(* IEC 61131-3 sources: daoli-st-library/DL_Device (part 4) *)

(* ---- FB_DL_PortDiagAggregator.st ---- *)
(*==============================================================================
 * 组件名称 (Component)  : FB_DL_PortDiagAggregator
 * 所属子库 (Sublibrary) : DL_Device
 * 当前版本 (Version)    : 1.0.0
 * 组件分类 (Category)   : 功能块（FUNCTION_BLOCK）· 设备诊断 · 端口级聚合仲裁
 * 兼容性   (Platform)   : CODESYS 3.5 / TwinCAT 3 / 汇川 InoProShop / Schneider
 *                         Machine Expert；仅位与运算、TON、R_TRIG 与标准类型
 * 功能描述 (Function)   : 把最多 8 个现场总线通讯端口的链路状态、诊断码、
 *                         CRC 错误累计计数聚合成单一故障掩码、首出端口号、
 *                         首出诊断码与错误风暴标志，解决「多端口同时报警时
 *                         HMI 只看到最后一条」的现场痛点。本块只做端口级
 *                         （通讯物理端口）聚合与首出仲裁，不做模块级位域解析。
 * 边界声明 (Boundary)   : FB_DL_AxiolineDiagLatch 负责本地总线模块级（槽号加
 *                         位域）诊断锁存；FB_DL_PdiReadScheduler 负责参数对象
 *                         读取调度；本块数据源是「端口计数与端口诊断码」，
 *                         三者数据源不同、码段不共享、互不可替。
 * 首出语义 (First-out)  : 仅在无锁存时仲裁，同拍多端口故障取端口号最小者
 *                         （低号端口更靠近主站，是现场排故的默认因果顺序）；
 *                         锁存后不再更新，只有复位上升沿可清。复位处理放在
 *                         仲裁之后，保证复位当拍首出即为空，下一拍重新仲裁。
 * 拍序纪律 (Cycle order) : 本块属监视型，但「窗口差分」有硬拍序：增量必须在
 *                         装载前算出并转出，否则窗口结束拍装载当拍增量恒为 0。
 *                         故输出数组先转出（上一段快照）后装载（下一段基准）。
 * 风暴语义 (Burst)      : 风暴是趋势事件，不锁存；eBurst 只停留一拍，该拍
 *                         置 bBurstDetected 单拍标志，供上层做趋势记录或
 *                         降低总线负载，不参与 bError 判定。
 * 开源溯源 (Origin)     : plcnext-community / profibus-diag / namur-ne107。参考
 *                         PLCnext 官方帮助与 PROFIBUS 诊断公开手册的端口诊断
 *                         功能分类与参数域（端口号、链路状态、诊断码、错误
 *                         计数器、错误风暴阈值），只借分类与参数域，端口数
 *                         上限、掩码位序、枚举、状态机、码位与全部算法 100%
 *                         自有，输入一律经引脚注入，不绑定任何厂商系统变量，
 *                         clean-room 实现，不构成衍生作品。
 * 依赖     (Depends)    : 无 DL_ 内部依赖；仅 Standard.library 的 TON / R_TRIG
 * 故障码表 (Error codes):
 *   16#0003_0140【信息级】端口数超上限已钳位（只进码与趋势，不置故障位）
 *   16#0003_0141【信息级】统计窗口参数越界已钳位（只进码，不置故障位）
 *   16#0003_0300【故障级】端口故障锁存（伴随故障掩码非零，置 bError）
 *   16#0003_0301【故障级】诊断源未注入（端口数小于 1，置 bError）
 *   16#0003_0307【故障级】非法状态兜底（置 bError）
 * 码位占用 (Slot)       : 信息级 0140 / 0141；故障级 0300 / 0301 / 0307。
 *                         全部落在 R11 本件分配块内，无跨块借用。
 * 写入点次序 (Write order) :
 *   ① ePhase   ：段 8 状态机（唯一位移点），段 10 复位分支可回 eIdle
 *   ② uErrorId ：段 11 单一优先级链（0307 优于 0301 优于 0300 优于 0141
 *                 优于 0140），全拍只写一次，杜绝多分支互相覆盖
 *   ③ 首出锁存 ：段 9 仲裁（仅未锁存时）→ 段 10 复位（唯一清除点）
 *   ④ 基准计数 ：段 8 窗口结束拍装载，段 5 只读，永不与增量同拍混用
 * 验收向量 (Acceptance) :
 *   V1 端口 2 与端口 5 故障，其余正常 → 故障掩码 16#0012、存在端口故障为真
 *   V2 端口 5 先故障、端口 2 后故障 → 首出端口 5；复位后才可更新为 2
 *   V3 窗口 1 秒、阈值 10、端口 3 计数 100 增至 115 → 窗口结束拍增量为 15、
 *      风暴标志单拍为真
 *   V4 端口 4 计数 16#FFFF_FFFF 回绕到 3 → 增量为 3，不出现巨大正数
 *   V5 端口数 12 → 钳位 8、码 16#0003_0140、bError 为假
 * 红线自检 (Redline)    : R1 零全局变量表与外部变量引用 ｜ R2 零物理地址直写
 *                         R3 纯 IEC 61131-3 ｜ R4 防除零、防越界、无浮点判等
 *                         R5 全变量中英双语同行注释 ｜ R6 ENUM 加 CASE 加 ELSE
 *                         R7 TON 与 R_TRIG 全部在 CASE 之外无条件刷新
 *                         R8 信息级码不置 bError，故障级码才置
 * 修订历史 (Revision)   :
 *   2026-11-15  v1.0.0  首版落盘（Round 11 · 泳道 B · T1-7 端口诊断族）
 *============================================================================*)

(*------------------------------------------------------------------------------
 * 枚举: E_DL_PortDiagPhase（本块相位，归属本功能块并同文件发布）
 *       Phase enumeration owned by this block and published in the same file
 *-----------------------------------------------------------------------------*)
TYPE E_DL_PortDiagPhase :
(
    eIdle    := 0,   // 待机：未使能或端口数非法，掩码清零、首出保持 / Idle, mask cleared, first-out kept
    eMonitor := 10,  // 监视：逐拍算增量、逐端口去抖、窗口边界拍评估 / Monitoring, deltas and debounce running
    eBurst   := 20,  // 风暴：仅停留一拍，置单拍风暴标志后回监视 / Burst, one cycle only then back to monitor
    eFault   := 99   // 故障：诊断源缺失或非法状态，需复位退出 / Fault, needs a reset to leave
);
END_TYPE

(*------------------------------------------------------------------------------
 * 结构体: ST_DL_PortDiagState（跨周期状态，由调用方持有）
 *         Persistent state structure, owned by the caller
 *         注意：本结构体是跨周期数据，E_DL_PortDiagPhase 是相位枚举，
 *         二者刻意同名不同前缀，禁止相互替换使用
 *-----------------------------------------------------------------------------*)
TYPE ST_DL_PortDiagState :
STRUCT
    auPrevCnt   : ARRAY[1..8] OF UDINT;  // 上窗口各端口 CRC 计数基准 [次] / Previous window CRC counter per port
    nLatchPort  : INT;                   // 首出故障端口号 [1..8]，0 表示无 / First-out port number, zero means none
    uLatchCode  : UDINT;                 // 首出端口诊断码 [代码]，0 表示无 / First-out diagnostic code, zero means none
    bLatchValid : BOOL;                  // 首出锁存有效，仅复位可清 [-] / First-out latch valid, reset clears it
END_STRUCT
END_TYPE

(*==============================================================================
 * 逐拍推演 (Cycle-by-cycle trace)：
 *   场景 A 双端口故障（端口 2 与端口 5）
 *     拍 k 段 6 逐端口判定为真并启动各自去抖；段 9 见无锁存，取最小号端口 2
 *          锁存端口 2 与端口 2 的诊断码；段 11 掩码为 16#0012、置 0300
 *   场景 B 首出不覆盖（端口 5 先、端口 2 后）
 *     拍 k 端口 5 故障，锁存 5；拍 k+n 端口 2 也故障，但 bLatchValid 已真，
 *          段 9 只观测不覆盖，首出维持 5；复位后下一拍重新仲裁得 2
 *   场景 C 错误风暴（窗口 1 秒、阈值 10、端口 3 计数 100 增到 115）
 *     窗口内段 5 每拍算 115 减 100 得增量 15；窗口结束拍段 8 评估 15 大于 10，
 *          转 eBurst；下一拍 eBurst 置风暴单拍标志，回 eMonitor，同时已装载
 *          新基准 115，故下一窗口增量从 0 起算
 *   场景 D 计数回绕（端口 4 由 16#FFFF_FFFF 变为 3）
 *     段 5 判出当前值小于基准，按归零处理取 3，绝不出现巨大正数假风暴
 *   场景 E 端口数超上限（端口数 12）
 *     段 3 钳位为 8 并标记；段 11 单独置 0140，bError 保持假
 *============================================================================*)

FUNCTION_BLOCK FB_DL_PortDiagAggregator
VAR_INPUT
    bEnable          : BOOL;                              // 使能，FALSE 时掩码清零、首出保持 [-] / Enable, clears mask, holds first-out
    bReset           : BOOL;                              // 复位首出锁存，上升沿有效 [-] / Reset the first-out latch on a rising edge
    nPortCount       : INT;                               // 实际端口数 [个]，有效域 1 到 8 / Port count, valid range one to eight
    abPortLinkOk     : ARRAY[1..8] OF BOOL;               // 各端口链路正常标志 [TRUE=正常] / Per-port link up flags
    auPortErrCode    : ARRAY[1..8] OF UDINT;              // 各端口诊断码 [代码]，0 表示正常 / Per-port diagnostic code, zero means OK
    auPortCrcErrCnt  : ARRAY[1..8] OF UDINT;              // 各端口 CRC 错误累计计数 [次] / Per-port CRC error counter
    nBurstThreshold  : UDINT := 10;                       // 窗口内错误增量阈值 [次]，0 表示不判风暴 / Burst threshold per window, zero disables
    tBurstWindow     : TIME := T#1S;                      // 错误风暴统计窗口长度 [毫秒] / Burst evaluation window
    tDebounce        : TIME := T#200MS;                   // 端口故障确认去抖时间 [毫秒]，0 表示不去抖 / Port fault debounce, zero disables
END_VAR
VAR_OUTPUT
    bAnyPortFault    : BOOL;                              // 任一端口故障，等价掩码非零 [-] / Any port faulted, mask is non-zero
    bBurstDetected   : BOOL;                              // 错误风暴单拍标志，仅 eBurst 拍为真 [-] / Burst single-scan flag, true only in the burst cycle
    uPortFaultMask   : WORD;                              // 端口故障掩码，位 n 对应端口 n 加一 [位串] / Port fault mask, bit n is port n plus one
    nFirstFaultPort  : INT;                               // 首出故障端口号 [1..8]，0 表示无 / First-fault port number, zero means none
    uFirstFaultCode  : UDINT;                             // 首出端口诊断码 [代码]，与端口号同拍锁存 / First-fault diagnostic code latched with the port
    auPortDelta      : ARRAY[1..8] OF UDINT;              // 本窗口各端口错误增量 [次] / Per-port error increment of this window
    eState           : E_DL_PortDiagPhase;                // 主状态机当前相位 [-] / Current phase of the main state machine
    bError           : BOOL;                              // 故障级锁存，仅 0300 0301 0307 置位 [-] / Latched fault, only fault level codes set it
    uErrorId         : UDINT;                             // 事件码，0 表示无事件 [代码] / Event code, zero means none
END_VAR
VAR_IN_OUT
    stState          : ST_DL_PortDiagState;               // 跨周期状态：基准计数与首出锁存 [-] / Persistent state, baseline counters and first-out latch
END_VAR
VAR
    fbTrigReset      : R_TRIG;                            // 复位沿检测，CASE 之外无条件刷新 [-] / Reset edge detector, refreshed outside the CASE
    fbTonWindow      : TON;                               // 风暴统计窗口计时，CASE 之外无条件刷新 / Burst window timer, refreshed outside the CASE
    afbDebounce      : ARRAY[1..8] OF TON;                // 逐端口故障去抖定时器组，循环内无条件全刷新 / Per-port debounce timers, all refreshed every cycle
    bInit            : BOOL := FALSE;                     // 首扫标志，初值 FALSE，判据 NOT bInit [-] / First-scan flag initialised FALSE
    ePhase           : E_DL_PortDiagPhase := E_DL_PortDiagPhase.eIdle;  // 内部相位，对外经 eState 输出 / Internal phase, exported as eState
    nPortClamped     : INT;                               // 钳位后的端口数 [个]，0 到 8 / Clamped port count, zero to eight
    tWinUse          : TIME;                              // 实际生效的窗口长度 [毫秒] / Effective window length
    tDebUse          : TIME;                              // 实际生效的去抖时间 [毫秒] / Effective debounce time
    bWinRun          : BOOL;                              // 窗口计时器输入，边界拍拉低以重启窗口 / Window timer input, dropped on the boundary cycle
    bWinElapsed      : BOOL;                              // 窗口结束拍标志 [-] / Window boundary flag
    abRawFault       : ARRAY[1..8] OF BOOL;               // 端口原始故障（未去抖）[-] / Raw per-port fault before debouncing
    uMaskBuild       : WORD;                              // 去抖后故障掩码装配中间量 [位串] / Fault mask under assembly after debounce
    auRawDelta       : ARRAY[1..8] OF UDINT;              // 本拍增量装配中间量 [次] / Increment under assembly of this cycle
    auOutDelta       : ARRAY[1..8] OF UDINT;              // 增量输出快照，先转出后装载 [-] / Increment snapshot exported before reloading the baseline
    uMaxDelta        : UDINT;                             // 窗口内最大增量 [次] / Maximum increment inside the window
    nFirstScanPort   : INT;                               // 仲裁临时：最小号故障端口 [1..8] / Arbitration temporary, lowest faulted port
    uFirstScanCode   : UDINT;                             // 仲裁临时：该端口诊断码 [代码] / Arbitration temporary, that port diagnostic code
    bPortCntClamped  : BOOL;                              // 端口数超上限被钳位的标记 [-] / Flag, port count was clamped
    bParamClamped    : BOOL;                              // 时间参数越界被钳位的标记 [-] / Flag, a time parameter was clamped
    bStateIllegal    : BOOL;                              // 非法状态被兜底捕获的标记 [-] / Flag, an illegal state was captured
    i                : INT;                               // 端口遍历索引 [1..8] / Port loop index
END_VAR
VAR CONSTANT
    DL_PORT_MAX      : INT := 8;                          // 端口上限 [个] / Maximum port count
    DL_PORT_MASK_ALL : WORD := 16#00FF;                   // 八端口全掩码 [位串] / All eight port mask
    DL_MASK_ONE      : WORD := 16#0001;                   // 单端口基准位 [位串] / Single port base bit
    DL_WIN_MIN       : TIME := T#1MS;                     // 窗口长度下限 [毫秒]，防 0 窗口 / Minimum window length, guards a zero window
    DL_DEB_MIN       : TIME := T#1MS;                     // 去抖时间下限 [毫秒]，非零时套用 / Minimum debounce when not disabled
    DL_TIME_ZERO     : TIME := T#0MS;                     // 时间零值基准 [毫秒] / Time zero reference
    DL_BURST_MARGIN  : UDINT := 0;                        // 增量比较余量 [次]，保留语义位 / Increment comparison margin, reserved semantic slot
END_VAR

(*------------------------------------------------------------------------------
 * 段 1｜沿检测无条件刷新（R7 红线：CASE 之外每拍必刷）
 *      Edge detection refreshed unconditionally outside the CASE
 *-----------------------------------------------------------------------------*)
fbTrigReset(CLK := bReset);

(*------------------------------------------------------------------------------
 * 段 2｜首扫初始化（R19 唯一合法范式：初值 FALSE，判据 NOT bInit）
 *      First-scan initialisation, the canonical R19 pattern
 *-----------------------------------------------------------------------------*)
IF NOT bInit THEN
    FOR i := 1 TO DL_PORT_MAX DO
        stState.auPrevCnt[i] := 0;               // 基准计数清零，避免首窗口假风暴
        auOutDelta[i]        := 0;               // 增量输出清零，HMI 初值确定
    END_FOR
    stState.nLatchPort     := 0;                 // 首出端口号：0 表示无
    stState.uLatchCode     := 0;                 // 首出诊断码：0 表示无
    stState.bLatchValid    := FALSE;             // 首出锁存无效
    ePhase                 := E_DL_PortDiagPhase.eIdle;
    nPortClamped           := 0;
    uMaskBuild             := 16#0000;
    bWinRun                := FALSE;
    bBurstDetected         := FALSE;
    bPortCntClamped        := FALSE;
    bParamClamped          := FALSE;
    bStateIllegal          := FALSE;
    eState                 := E_DL_PortDiagPhase.eIdle;
    uErrorId               := 16#0000_0000;
    bError                 := FALSE;
    bInit                  := TRUE;              // 首扫只做一次
END_IF

(*------------------------------------------------------------------------------
 * 段 3｜端口数钳位（越界只钳位，不越界访问数组）
 *      Port count clamping, never index outside the array
 *-----------------------------------------------------------------------------*)
bPortCntClamped := FALSE;                        // 本拍标记预清零，避免历史残留
IF nPortCount < 1 THEN
    nPortClamped := 0;                           // 无诊断源：交由状态机转故障
ELSIF nPortCount > DL_PORT_MAX THEN
    nPortClamped    := DL_PORT_MAX;              // 超上限钳位到 8
    bPortCntClamped := TRUE;                     // 标记待置信息级码 0140
ELSE
    nPortClamped := nPortCount;
END_IF

(*------------------------------------------------------------------------------
 * 段 4｜时间参数钳位（0 有明确语义，不得与越界混为一谈）
 *      Time parameter clamping, zero keeps its documented meaning
 *-----------------------------------------------------------------------------*)
bParamClamped := FALSE;                          // 本拍标记预清零，避免历史残留
IF tBurstWindow <= DL_TIME_ZERO THEN
    tWinUse      := DL_WIN_MIN;                  // 0 窗口会让计时器每拍立即到期
    bParamClamped := TRUE;
ELSIF tBurstWindow < DL_WIN_MIN THEN
    tWinUse      := DL_WIN_MIN;
    bParamClamped := TRUE;
ELSE
    tWinUse := tBurstWindow;
END_IF

IF tDebounce < DL_TIME_ZERO THEN
    tDebUse      := DL_DEB_MIN;                  // 负时间不可能，按最小值兜底
    bParamClamped := TRUE;
ELSE
    tDebUse := tDebounce;                        // 0 表示不去抖，原样透传
END_IF

(*------------------------------------------------------------------------------
 * 段 5｜增量差分（回绕按归零处理，UDINT 语义不产生负数）
 *      Increment differencing, a wrapped counter is treated as a restart
 *      纪律：本段只读基准，装载基准只在段 8 窗口结束拍执行
 *-----------------------------------------------------------------------------*)
FOR i := 1 TO DL_PORT_MAX DO
    IF i > nPortClamped THEN
        auRawDelta[i] := 0;                      // 超出实际端口数一律记为 0
        auOutDelta[i] := 0;
    ELSIF auPortCrcErrCnt[i] < stState.auPrevCnt[i] THEN
        auRawDelta[i] := auPortCrcErrCnt[i];     // 计数器回绕或复位：按归零处理
        auOutDelta[i] := auRawDelta[i];
    ELSE
        auRawDelta[i] := auPortCrcErrCnt[i] - stState.auPrevCnt[i];
        auOutDelta[i] := auRawDelta[i];          // 先转出快照，供段 11 输出
    END_IF
END_FOR

(*------------------------------------------------------------------------------
 * 段 6｜端口故障判定与逐端口去抖（掩码装配）
 *      Per-port fault evaluation with per-port debounce and mask assembly
 *      定时器组在循环内对全部八端口无条件刷新，不因端口数少而漏刷
 *-----------------------------------------------------------------------------*)
uMaskBuild := 16#0000;
FOR i := 1 TO DL_PORT_MAX DO
    IF bEnable AND (i <= nPortClamped) AND ((NOT abPortLinkOk[i]) OR (auPortErrCode[i] <> UDINT#0)) THEN
        abRawFault[i] := TRUE;                   // 链路断或诊断码非零即原始故障
    ELSE
        abRawFault[i] := FALSE;
    END_IF
    afbDebounce[i](IN := abRawFault[i], PT := tDebUse);
    IF afbDebounce[i].Q THEN
        uMaskBuild := uMaskBuild OR SHL(DL_MASK_ONE, i - 1);  // 去抖成立才进位
    END_IF
END_FOR

(*------------------------------------------------------------------------------
 * 段 7｜窗口计时（无条件刷新，输入取自上一拍的运行允许位）
 *      Window timer refreshed unconditionally, input from the previous cycle
 *-----------------------------------------------------------------------------*)
fbTonWindow(IN := bWinRun, PT := tWinUse);
bWinElapsed := fbTonWindow.Q;

(*------------------------------------------------------------------------------
 * 段 8｜主状态机（ENUM 加 CASE，含 ELSE 兜底；每成员均有对应标签）
 *      Main state machine, one label per enumeration member plus a fallback
 *-----------------------------------------------------------------------------*)
bBurstDetected := FALSE;                         // 单拍标志预清零：只在 eBurst 拍置真
CASE ePhase OF
    E_DL_PortDiagPhase.eIdle:
        bWinRun := FALSE;                        // 待机不跑窗口，避免脏计时
        IF bEnable AND (nPortClamped >= 1) THEN
            ePhase  := E_DL_PortDiagPhase.eMonitor;
            bWinRun := TRUE;                     // 进入监视即启动首个窗口
        ELSIF bEnable AND (nPortClamped < 1) THEN
            ePhase := E_DL_PortDiagPhase.eFault; // 诊断源未注入：故障级 0301
        END_IF

    E_DL_PortDiagPhase.eMonitor:
        IF NOT bEnable THEN
            ePhase     := E_DL_PortDiagPhase.eIdle;
            bWinRun    := FALSE;
            uMaskBuild := 16#0000;               // 未使能掩码清零，首出保持
        ELSIF nPortClamped < 1 THEN
            ePhase  := E_DL_PortDiagPhase.eFault;
            bWinRun := FALSE;
        ELSIF bWinElapsed THEN
            uMaxDelta     := 0;                  // 窗口结束拍：求最大增量
            FOR i := 1 TO nPortClamped DO
                IF auRawDelta[i] > uMaxDelta THEN
                    uMaxDelta := auRawDelta[i];
                END_IF
            END_FOR
            IF (nBurstThreshold > UDINT#0) AND (uMaxDelta > (nBurstThreshold + DL_BURST_MARGIN)) THEN
                ePhase := E_DL_PortDiagPhase.eBurst;   // 超阈值：下一拍置单拍标志
            ELSE
                ePhase := E_DL_PortDiagPhase.eMonitor; // 未超阈值：原地自保持
            END_IF
            FOR i := 1 TO DL_PORT_MAX DO
                stState.auPrevCnt[i] := auPortCrcErrCnt[i];  // 装载新基准
            END_FOR
            bWinRun := FALSE;                    // 拉低一拍，强制窗口重新起算
        ELSE
            bWinRun := TRUE;                     // 窗口内持续计时
        END_IF

    E_DL_PortDiagPhase.eBurst:
        bBurstDetected := TRUE;                  // 仅此一拍为真，不锁存，不进故障
        bWinRun        := FALSE;                 // 风暴拍不重启窗口，下一拍再说
        ePhase         := E_DL_PortDiagPhase.eMonitor;

    E_DL_PortDiagPhase.eFault:
        uMaskBuild := 16#0000;                   // 故障态不外送掩码，防误联锁
        bWinRun    := FALSE;
        IF NOT bEnable THEN
            ePhase := E_DL_PortDiagPhase.eIdle;  // 停使能可直接退出故障态
        END_IF

    ELSE
        ePhase        := E_DL_PortDiagPhase.eFault;   // 非法值兜底
        uMaskBuild    := 16#0000;
        bWinRun       := FALSE;
        bStateIllegal := TRUE;                   // 由段 11 统一置 0307
END_CASE

(*------------------------------------------------------------------------------
 * 段 9｜首出仲裁（仅未锁存时执行；升序取最小号端口，先到先得）
 *      First-out arbitration, only when not yet latched, lowest port wins
 *-----------------------------------------------------------------------------*)
IF (NOT stState.bLatchValid) AND uMaskBuild <> 16#0000 THEN
    nFirstScanPort := 0;
    uFirstScanCode := 0;
    FOR i := 1 TO nPortClamped DO
        IF ((uMaskBuild AND SHL(DL_MASK_ONE, i - 1)) <> 16#0000) AND (nFirstScanPort = 0) THEN
            nFirstScanPort := i;                       // 升序首个命中即最小号端口
            uFirstScanCode := auPortErrCode[i];
        END_IF
    END_FOR
    IF nFirstScanPort > 0 THEN
        stState.nLatchPort  := nFirstScanPort;
        stState.uLatchCode  := uFirstScanCode;
        stState.bLatchValid := TRUE;                   // 锁存后本窗口不再改写
    END_IF
END_IF

(*------------------------------------------------------------------------------
 * 段 10｜复位（放在仲裁之后，保证复位当拍首出即为空）
 *      Reset placed after arbitration so the first-out is empty this cycle
 *-----------------------------------------------------------------------------*)
IF fbTrigReset.Q THEN
    stState.nLatchPort  := 0;
    stState.uLatchCode  := 0;
    stState.bLatchValid := FALSE;
    bError              := FALSE;
    bStateIllegal       := FALSE;
    ePhase              := E_DL_PortDiagPhase.eIdle;   // 复位后回待机，再按使能重入
    bWinRun             := FALSE;
END_IF

(*------------------------------------------------------------------------------
 * 段 11｜输出归并与码位定级（单一优先级链，全拍只写一次 uErrorId）
 *      Output merge and single-priority error code resolution
 *-----------------------------------------------------------------------------*)
uPortFaultMask  := uMaskBuild AND DL_PORT_MASK_ALL;    // 屏蔽高位脏数据
bAnyPortFault   := (uPortFaultMask <> 16#0000);
nFirstFaultPort := stState.nLatchPort;
uFirstFaultCode := stState.uLatchCode;

IF bStateIllegal THEN
    uErrorId := 16#0003_0307;                          // 优先级一：非法状态
ELSIF (nPortClamped < 1) AND bEnable THEN
    uErrorId := 16#0003_0301;                          // 优先级二：诊断源缺失
ELSIF uPortFaultMask <> 16#0000 THEN
    uErrorId := 16#0003_0300;                          // 优先级三：端口故障锁存
ELSIF bParamClamped THEN
    uErrorId := 16#0003_0141;                          // 信息级：参数越界已钳位
ELSIF bPortCntClamped THEN
    uErrorId := 16#0003_0140;                          // 信息级：端口数越界已钳位
ELSE
    uErrorId := 16#0000_0000;
END_IF

(* 故障位只反映故障级：信息级码 0140 与 0141 绝不置故障位（R21） *)
bError := bStateIllegal
          OR ((nPortClamped < 1) AND bEnable)
          OR (uPortFaultMask <> 16#0000);

eState          := ePhase;                             // 相位每拍重写，供 HMI 诊断
auPortDelta[1]  := auOutDelta[1];                      // 增量数组逐元素转出，避免整数组赋值
auPortDelta[2]  := auOutDelta[2];
auPortDelta[3]  := auOutDelta[3];
auPortDelta[4]  := auOutDelta[4];
auPortDelta[5]  := auOutDelta[5];
auPortDelta[6]  := auOutDelta[6];
auPortDelta[7]  := auOutDelta[7];
auPortDelta[8]  := auOutDelta[8];
END_FUNCTION_BLOCK

(* ---- FB_DL_PortDiagBoard.st ---- *)
(*==============================================================================
 * 组件名称 (Component)  : FB_DL_PortDiagBoard
 * 所属子库 (Sublibrary) : DL_Device
 * 当前版本 (Version)    : 1.0.0
 * 组件分类 (Category)   : 功能块（FUNCTION_BLOCK）· 设备诊断 · 多组端口看板与首出仲裁
 * 兼容性   (Platform)   : CODESYS 3.5 / TwinCAT 3 / 汇川 InoProShop / Schneider
 *                         Machine Expert；纯 IEC 61131-3（第 3 版）语法，
 *                         仅依赖 Standard.library（R_TRIG），零厂商方言
 * 功能描述 (Function)   : 把最多 4 个端口诊断聚合组（每组最多 8 端口）汇总为一张看板：
 *                         屏蔽超界位后的各组掩码、全局故障端口总数、全局首出端口
 *                         （组号加端口号加诊断码），以及按「组号优先、端口号次之」稳定
 *                         排序的前 3 个待修端口。回答现场两个问题：现在还剩几个端口坏、
 *                         先修哪一个。
 * 分层声明 (Layering)   : ① 本件是「汇总层」，只消费端口级聚合结果（掩码加组内首出
 *                         码），不实例化上游聚合块、不重算端口明细——聚合器实例由调用方
 *                         按组各自持有，重复实例化会造成同一批端口被算两遍；
 *                         ② 不读模块级状态字（模块级归本地总线诊断锁存件，端口级归聚合
 *                         器，参数对象级归参数回读调度件，三层数据源分账已在 R11 收口）；
 *                         ③ 不绑定任何总线驱动，全部数据经引脚注入。
 * 职责边界 (Scope)      : 不做端口去抖（聚合器职责）、不做报警确认与搁置、不做历史趋势
 *                         归档、不做跨机架分组切换（组数运行期变化按钳位处理）。
 * 组数语义 (Grouping)   : 组是「同一块远程 IO 卡或同一台交换机的 8 个端口」的物理分组，
 *                         组号小者更靠近主站，故首出仲裁取组号最小、再取端口号最小，
 *                         这与现场排故的因果顺序一致。
 * 开源溯源 (Origin)     : 来源标签 plcnext-diag 加 roadmap-p0。原创实现（参考 T1-7
 *                         PLCnext 端口诊断四元组的分类与参数域，以及 ROADMAP §15.3 P0
 *                         条目的「看板加首出」需求定义）。仅借分类层次、参数域与验收
 *                         口径，掩码位序、首出三律、Top 排序编码、枚举、状态机与全部
 *                         码位 100% 本库独立设计，clean-room 实现，零代码行复制。
 *                         PLCnext 帮助文档为厂商公开资料，此处按最严口径「只借结构与
 *                         参数域」处置，不构成衍生作品。
 * 依赖     (Depends)    : 无 DL_ 内部依赖；Standard.library: R_TRIG
 * 故障码表 (Error codes):
 *   16#0003_0149【信息级】组数超上限已钳位到 4（只影响显示范围，不置故障位）
 *   16#0003_014A【信息级】某组端口数超上限已钳位到 8（组态常见，非错误）
 *   16#0003_014B【信息级】掩码超界位已屏蔽（绝不把不存在的端口计入故障数）
 *   16#0003_014C【信息级】组内声明首出端口与掩码推导值不一致（数据源未同步）
 *   16#0003_030B【故障段趋势码】单拍掩码变化位数超阈值，判为组态刷新；按规格
 *                         第 3.13 节「仅提示不锁存」处置：只透出一拍，不置故障位
 *   16#0003_0309【故障级】组数小于 1，无诊断源（锁存，置故障位）
 *   16#0003_030A【故障级】某组端口数小于 1，该组掩码含义不可信（锁存，置故障位）
 *   16#0003_030C【故障级】非法状态兜底（锁存，置故障位，终端安全态）
 * 码位占用 (Slot)       : 信息级 0149 / 014A / 014B / 014C；故障级 0309 / 030A / 030B / 030C。
 *                         全部落在 R12 本件分配块内，无跨块借用、无段外哨兵值。
 * 拍序纪律 (Cycle order) :
 *   ① ePhase      ：段 4 状态机（唯一位移点），段 6 复位分支是唯一回退点
 *   ② 首出锁存    ：段 4 的 eScanning 分支（仅未锁存时仲裁）→ 段 5 换出 → 段 6 复位清除
 *   ③ 输出码      ：段 7 单一优先级链，全拍只写一次 uErrorId，杜绝多分支互相覆盖
 *   ④ 掩码基准    ：段 4 的 eScanning 分支末尾装载，与风暴判定同段且判在读后写前
 * 首出三律 (First-out)  : ① 仅在无锁存时仲裁；② 同拍多端口故障取组号最小、再取端口号
 *                         最小；③ 复位在仲裁之后执行，故复位当拍首出为空、下一拍重新
 *                         仲裁（与 R11 端口聚合器同口径）。
 * 验收向量 (Acceptance) :
 *   V1 单组超界位：组数 1、端口数 8、掩码 16#0101 → 位 8 对应端口 9 超界被屏蔽，
 *      掩码出 16#0001、总故障 1、首出 1 组 1 号、码 014B
 *   V2 双组排序：两组端口数 8，掩码 16#0004 与 16#0003 → 总数 3、首出 1 组 3 号、
 *      待修序 13、21、22（编码为组号乘 10 加端口号）
 *   V3 复位时序：与 V2 同参，复位上升沿当拍首出为空，下一拍重新仲裁回 1 组 3 号
 *   V4 无诊断源：组数 0 → 钳为 1、故障位置位、码 0309
 *   V5 空组：第 1 组端口数 0 → 钳为 1、故障位置位、码 030A
 * 偏离留档 (Deviation)  :
 *   ① 规格第 3.13 节算法要点对「端口数超上限」写 014A、对「端口数越界」的边界说明
 *      又写 030A。本件按语义拆分：大于 8 属组态多填，按信息级 014A 只钳位；小于 1
 *      属无有效端口（掩码含义不可信），按故障级 030A 锁存——与验收向量 V5 完全一致。
 *   ② 规格未给 anGroupFirstPort 的用途。本件把它用作「声明值与掩码推导值」的一致性
 *      校验（为 0 视为未填、不校验），不一致只置信息级 014C，避免该引脚悬空无意义。
 *   ③ 030B 落在故障段但不置故障位，理由见上方故障码表，属规格原文要求的「仅提示不
 *      锁存」，不是定级笔误。
 * 修订历史 (Revision)   :
 *   2026-11-15  v1.0.0  首版落盘（R12 · 泳道 C · 端口诊断看板 P0 件）
 *============================================================================*)

(*------------------------------------------------------------------------------
 * 枚举: E_DL_BoardPhase（本块相位，归属本功能块并同文件发布）
 *       Phase enumeration owned by this block and published in the same file
 *-----------------------------------------------------------------------------*)
TYPE E_DL_BoardPhase :
(
    eIdle     := 0,   // 待机：钳位参数后即转扫描，或未使能时清掩码保首出 / Idle, clamps parameters then moves on to scanning
    eScanning := 10,  // 扫描：一趟完成屏蔽、计数、首出仲裁与待修排序，本拍结束回待机 / Scanning, the whole sweep completes in one pass
    eFault    := 99   // 故障：无诊断源、空组或非法状态，需复位退出 / Fault, needs a reset to leave
);
END_TYPE

(*------------------------------------------------------------------------------
 * 结构体: ST_DL_BoardState（跨周期状态，由调用方持有）
 *         Persistent state structure, owned by the caller
 *         说明：首出锁存是「诊断证据」，掉使能不清、只有复位沿才清；
 *               anLastMask 用于掩码跳变风暴的差分基准
 *-----------------------------------------------------------------------------*)
TYPE ST_DL_BoardState :
STRUCT
    nLatchedGroup : INT;                     // 首出锁存组号 [1..4]，0 表示无 / Latched first-out group, zero means none
    nLatchedPort  : INT;                     // 首出锁存端口号 [1..8]，0 表示无 / Latched first-out port, zero means none
    uLatchedCode  : UDINT;                   // 首出锁存诊断码 [代码]，0 表示未填 / Latched first-out diagnostic code, zero means not filled
    bLatchValid   : BOOL;                    // 首出锁存有效，仅复位沿可清 / First-out latch valid, cleared by the reset edge only
    anLastMask    : ARRAY[1..4] OF WORD;     // 上次各组掩码快照，用于跳变风暴差分 [位串] / Previous per-group mask for burst differencing
END_STRUCT
END_TYPE

FUNCTION_BLOCK FB_DL_PortDiagBoard
VAR_INPUT
    bEnable          : BOOL;                              // 看板使能，FALSE 时掩码清零而首出保持 [-] / Enable, masks are cleared while the first-out latch is kept
    bReset           : BOOL;                              // 复位首出锁存，上升沿有效 [-] / Rising edge clears the first-out latch
    nGroupCount      : INT := 1;                          // 聚合组数 [组]，有效域 1 到 4 / Group count, valid range one to four
    anGroupFaultMask : ARRAY[1..4] OF WORD;               // 各组端口故障掩码，位 n 减一 对应端口 n [位串] / Per-group fault mask, bit n minus one is port n
    anGroupPortCount : ARRAY[1..4] OF INT;                // 各组实际端口数 [个]，有效域 1 到 8 / Ports per group, valid range one to eight
    anGroupFirstPort : ARRAY[1..4] OF INT;                // 各组声明首出端口号，0 表示未填不校验 [端口号] / Declared first-out port, zero skips the cross check
    auGroupFirstCode : ARRAY[1..4] OF UDINT;              // 各组组内首出诊断码 [代码]，0 表示未填 / Per-group first-out diagnostic code, zero means not filled
END_VAR
VAR_OUTPUT
    nTotalFaultPort  : INT;                               // 全局故障端口总数 [个] / Total faulted ports across the enabled groups
    nFirstGroup      : INT;                               // 全局首出组号 [1..4]，0 表示无 / Global first-out group, zero means none
    nFirstPort       : INT;                               // 全局首出端口号 [1..8]，0 表示无 / Global first-out port, zero means none
    uFirstCode       : UDINT;                             // 全局首出诊断码 [代码]，0 表示未填 / Global first-out diagnostic code
    anGroupMaskOut   : ARRAY[1..4] OF WORD;               // 屏蔽超界位后的各组掩码 [位串] / Sanitised per-group masks
    anTopPortNo      : ARRAY[1..3] OF INT;                // 待修端口编码，组号乘 10 加端口号，0 表示空位 [编码] / Top repair ports encoded as group times ten plus port
    auTopPortCode    : ARRAY[1..3] OF UDINT;              // 待修端口对应诊断码 [代码] / Diagnostic code of each top repair port
    bAnyFault        : BOOL;                              // 总故障数大于 0 [-] / Any faulted port present
    bError           : BOOL;                              // 故障级锁存，仅 0309 030A 030C 置位 [-] / Latched fault, only fault level codes set it
    uErrorId         : UDINT;                             // 事件码，0 表示无事件 [代码] / Event code, zero means none
    eState           : E_DL_BoardPhase;                   // 主状态机当前相位 [-] / Current phase of the main state machine
END_VAR
VAR_IN_OUT
    stBoard          : ST_DL_BoardState;                  // 跨周期：首出锁存与掩码差分基准 [-] / Persistent first-out latch and mask baseline
END_VAR
VAR
    fbTrigReset      : R_TRIG;                            // 复位沿检测，主周期无条件刷新 [-] / Reset edge detector, refreshed unconditionally
    ePhase           : E_DL_BoardPhase := E_DL_BoardPhase.eIdle; // 内部相位，对外经 eState 输出 [-] / Internal phase exported as eState
    bInit            : BOOL := FALSE;                     // 首扫标志，初值 FALSE，判据取非 [-] / First-scan flag initialised FALSE
    bMaskBase        : BOOL := FALSE;                     // 掩码差分基准已装载 [-] / Mask baseline loaded flag
    bFaultLatch      : BOOL;                              // 故障锁存，仅复位分支清除 [-] / Fault latch, cleared by the reset path only
    uErrInt          : UDINT;                             // 故障级码寄存，锁存型 [代码] / Latched fault level code register
    uInfoCode        : UDINT;                             // 本拍信息级码，每拍重算 [代码] / Info level code recomputed every scan
    nGroupUse        : INT;                               // 生效组数，钳位后 [组] / Effective group count after clamping
    auPortCntUse     : ARRAY[1..4] OF INT;                // 生效端口数，钳位后 [个] / Effective port count per group after clamping
    uBuildMask       : WORD;                              // 掩码装配中间量 [位串] / Mask under assembly
    uDiff            : WORD;                              // 掩码差分中间量 [位串] / Mask difference under evaluation
    nTotal           : INT;                               // 故障端口累加计数 [个] / Faulted port counter
    nMinPort         : INT;                               // 组内最小故障端口号 [1..8]，0 表示无 / Lowest faulted port inside a group
    nBitScan         : INT;                               // 掩码跳变位计数 [位] / Changed bit counter for the burst check
    nScanGroup       : INT;                               // 仲裁扫描组号 [1..4] / Arbitration group index
    nScanPort        : INT;                               // 仲裁扫描端口号 [1..8] / Arbitration port index
    bFound           : BOOL;                              // 仲裁命中标志 [-] / Arbitration hit flag
    nTopCount        : INT;                               // 已填待修位个数 [个] / Filled top repair slots
    nGuard           : DINT;                              // 循环守卫计数 [次]，上限常量化 / Loop guard counter with a constant bound
    bMaskClamped     : BOOL;                              // 本拍存在掩码超界位被屏蔽 [-] / Mask bits were suppressed this scan
    bPortClamped     : BOOL;                              // 本拍存在端口数超上限被钳位 [-] / A port count was clamped this scan
    bGroupClamped    : BOOL;                              // 本拍组数超上限被钳位 [-] / The group count was clamped this scan
    bPortShort       : BOOL;                              // 本拍存在某组端口数小于 1 [-] / A group has no usable port this scan
    bGroupShort      : BOOL;                              // 本拍组数小于 1 [-] / The group count is below one this scan
    bPortDeclMismatch: BOOL;                              // 声明首出端口与推导值不一致 [-] / Declared first-out port differs from the derived one
    bMaskJump        : BOOL;                              // 单拍掩码跳变位超阈值 [-] / Mask changed in more bits than the threshold
    g                : INT;                               // 组循环索引 [1..4] / Group loop index
    p                : INT;                               // 端口循环索引 [1..8] / Port loop index
END_VAR
VAR CONSTANT
    DL_GROUP_MAX     : INT := 4;                          // 聚合组数上限 [组] / Maximum group count
    DL_PORT_MAX      : INT := 8;                          // 组内端口数上限 [个] / Maximum ports per group
    DL_TOP_N         : INT := 3;                          // 待修输出位个数 [个] / Number of top repair slots
    DL_GROUP_STRIDE  : INT := 10;                         // 端口编码步长，组号乘该值加端口号 / Encoding stride of the top repair code
    DL_JUMP_MAX      : INT := 8;                          // 单拍掩码跳变位阈值 [位] / Changed bit threshold per scan
    DL_GUARD_MAX     : DINT := 96;                        // 循环守卫上限 [次] / Loop guard bound
    DL_WORD_BITS     : INT := 16;                         // 掩码字宽，超界位屏蔽的遍历上限 [位] / Mask word width
    DL_MASK_ONE      : WORD := 16#0001;                   // 单端口基准位 [位串] / Single port base bit
    DL_MASK_NONE     : WORD := 16#0000;                   // 全零掩码基准 [位串] / All zero mask reference
END_VAR

(*------------------------------------------------------------------------------
 * 段 1｜输出确定性默认值（公约：出口先赋；单拍标志每拍预清零，R25 第一律）
 *      Deterministic defaults first, one-scan flags pre-cleared every scan
 *-----------------------------------------------------------------------------*)
bAnyFault         := FALSE;                     // 看板派生量预清零（Dashboard flag pre-cleared）
uInfoCode         := 16#0000_0000;              // 信息级码每拍重算（Info code recomputed every scan）
bMaskClamped      := FALSE;                     // 掩码屏蔽标记预清零（Mask suppression flag pre-cleared）
bPortClamped      := FALSE;                     // 端口数钳位标记预清零（Port clamp flag pre-cleared）
bGroupClamped     := FALSE;                     // 组数钳位标记预清零（Group clamp flag pre-cleared）
bPortShort        := FALSE;                     // 空组标记预清零（Empty group flag pre-cleared）
bGroupShort       := FALSE;                     // 无组标记预清零（No group flag pre-cleared）
bPortDeclMismatch := FALSE;                     // 声明一致性标记预清零（Declared mismatch flag pre-cleared）
bMaskJump         := FALSE;                     // 掩码跳变标记预清零（Mask jump flag pre-cleared）
nGuard            := 0;                         // 循环守卫清零（Loop guard cleared）

(*------------------------------------------------------------------------------
 * 段 2｜沿检测无条件刷新（红线：实例在 CASE 之外每拍必刷）
 *      Edge detection refreshed unconditionally outside the CASE
 *-----------------------------------------------------------------------------*)
fbTrigReset(CLK := bReset);

(*------------------------------------------------------------------------------
 * 段 3｜首扫初始化（唯一合法范式：初值 FALSE，判据取非）
 *      First-scan initialisation following the single legal pattern
 *-----------------------------------------------------------------------------*)
IF NOT bInit THEN
    FOR g := 1 TO DL_GROUP_MAX DO
        stBoard.anLastMask[g] := DL_MASK_NONE;  // 掩码差分基准清零，避免首拍假风暴（Baseline cleared to suppress a false burst）
        anGroupMaskOut[g]     := DL_MASK_NONE;  // 掩码出口清零，HMI 初值确定（Mask outlet cleared for a deterministic HMI start value）
    END_FOR
    FOR p := 1 TO DL_TOP_N DO
        anTopPortNo[p]   := 0;                  // 待修端口空位（Top repair slot empty）
        auTopPortCode[p] := 0;                  // 待修诊断码清零（Top repair code cleared）
    END_FOR
    stBoard.nLatchedGroup := 0;                 // 首出组号：0 表示无（No first-out group）
    stBoard.nLatchedPort  := 0;                 // 首出端口号：0 表示无（No first-out port）
    stBoard.uLatchedCode  := 0;                 // 首出码：0 表示未填（No first-out code）
    stBoard.bLatchValid   := FALSE;             // 首出锁存无效（First-out latch invalid）
    nTotalFaultPort       := 0;                 // 故障总数清零（Fault total cleared）
    nFirstGroup           := 0;                 // 首出组号出口清零（First-out group outlet cleared）
    nFirstPort            := 0;                 // 首出端口出口清零（First-out port outlet cleared）
    uFirstCode            := 0;                 // 首出码出口清零（First-out code outlet cleared）
    bFaultLatch           := FALSE;             // 故障锁存清零（Fault latch cleared）
    uErrInt               := 16#0000_0000;      // 故障码清零（Fault code cleared）
    bMaskBase             := FALSE;             // 差分基准待本拍装载（Baseline to be loaded this scan）
    ePhase                := E_DL_BoardPhase.eIdle; // 相位复位为待机（Phase reset to idle）
    bInit                 := TRUE;              // 首扫只做一次（First scan runs once）
END_IF

(*------------------------------------------------------------------------------
 * 段 4｜主状态机（枚举每个成员均有标签，末尾 ELSE 兜底到终端安全态）
 *      Main state machine, one label per member plus a trailing ELSE fallback
 *-----------------------------------------------------------------------------*)
CASE ePhase OF

    E_DL_BoardPhase.eIdle: // 待机：未使能则清掩码保首出，使能则钳位参数后转扫描
        IF NOT bEnable THEN
            FOR g := 1 TO DL_GROUP_MAX DO
                anGroupMaskOut[g] := DL_MASK_NONE;  // 掉使能掩码清零，防止下游误联锁（Masks cleared while disabled）
            END_FOR
            nTotalFaultPort := 0;               // 故障总数清零（Fault total cleared）
            bAnyFault       := FALSE;           // 无故障派生量（No fault derived）
            ePhase          := E_DL_BoardPhase.eIdle; // 保持在待机（Stay idle）
        ELSE
            IF nGroupCount < 1 THEN
                nGroupUse    := 1;              // 无组：先给 1 供后续诊断（Fall back to one group）
                bGroupShort  := TRUE;           // 标记待置 0309（Flag for code 0309）
            ELSIF nGroupCount > DL_GROUP_MAX THEN
                nGroupUse    := DL_GROUP_MAX;   // 超上限钳位（Clamp to the upper bound）
                bGroupClamped := TRUE;          // 标记待置 0149（Flag for code 0149）
            ELSE
                nGroupUse := nGroupCount;       // 合法组数直通（Valid group count passed through）
            END_IF
            FOR g := 1 TO DL_GROUP_MAX DO
                nGuard := nGuard + 1;           // 守卫递增（Guard incremented）
                IF nGuard > DL_GUARD_MAX THEN
                    EXIT;                       // 守卫到顶即退出，防死循环（Bail out at the guard bound）
                END_IF
                IF g <= nGroupUse THEN
                    IF anGroupPortCount[g] < 1 THEN
                        auPortCntUse[g] := 1;   // 空组：先给 1 供后续诊断（Empty group falls back to one port）
                        bPortShort      := TRUE; // 标记待置 030A（Flag for code 030A）
                    ELSIF anGroupPortCount[g] > DL_PORT_MAX THEN
                        auPortCntUse[g] := DL_PORT_MAX; // 超上限钳位（Clamp to the upper bound）
                        bPortClamped    := TRUE;        // 标记待置 014A（Flag for code 014A）
                    ELSE
                        auPortCntUse[g] := anGroupPortCount[g]; // 合法端口数直通（Valid port count passed through）
                    END_IF
                ELSE
                    auPortCntUse[g] := 0;       // 未启用组记 0，不参与扫描（Unused group marked zero）
                END_IF
            END_FOR
            IF bGroupShort THEN
                bFaultLatch := TRUE;                        // 无诊断源：锁故障（No diagnostic source, latch a fault）
                uErrInt     := 16#0003_0309;                // 0309 组数小于 1（Group count below one）
                ePhase      := E_DL_BoardPhase.eFault;      // 进故障态（Enter the fault state）
            ELSIF bPortShort THEN
                bFaultLatch := TRUE;                        // 空组：锁故障（Empty group latches a fault）
                uErrInt     := 16#0003_030A;                // 030A 端口数小于 1（Port count below one）
                ePhase      := E_DL_BoardPhase.eFault;      // 进故障态（Enter the fault state）
            ELSE
                ePhase := E_DL_BoardPhase.eScanning;        // 参数可用，进入扫描（Parameters usable, start scanning）
            END_IF
        END_IF

    E_DL_BoardPhase.eScanning: // 扫描：屏蔽、计数、首出仲裁、待修排序、跳变差分，一趟完成
        nTotal    := 0;                         // 故障计数清零（Fault counter cleared）
        nBitScan  := 0;                         // 跳变位计数清零（Changed bit counter cleared）
        (* ① 屏蔽超界位并统计故障数，同时取组内最小故障端口号 *)
        nGuard := 0;                            // 子段守卫清零（Guard reset for this pass）
        FOR g := 1 TO DL_GROUP_MAX DO
            nGuard := nGuard + 1;               // 守卫递增（Guard incremented）
            IF nGuard > DL_GUARD_MAX THEN
                EXIT;                           // 守卫到顶即退出（Bail out at the guard bound）
            END_IF
            IF g <= nGroupUse THEN
                uBuildMask := anGroupFaultMask[g];      // 取原始掩码（Take the raw mask）
                nMinPort   := 0;                        // 组内最小端口号预清零（Lowest port pre-cleared）
                FOR p := 1 TO DL_WORD_BITS DO
                    nGuard := nGuard + 1;               // 守卫递增（Guard incremented）
                    IF nGuard > DL_GUARD_MAX THEN
                        EXIT;                           // 守卫到顶即退出（Bail out at the guard bound）
                    END_IF
                    IF p > auPortCntUse[g] THEN
                        IF (uBuildMask AND SHL(DL_MASK_ONE, p - 1)) <> DL_MASK_NONE THEN
                            bMaskClamped := TRUE;       // 超界位有值：标记待置 014B（Out-of-range bit held a value）
                        END_IF
                        uBuildMask := uBuildMask AND (NOT SHL(DL_MASK_ONE, p - 1)); // 超界位清零（Clear the out-of-range bit）
                    ELSE
                        IF (uBuildMask AND SHL(DL_MASK_ONE, p - 1)) <> DL_MASK_NONE THEN
                            nTotal := nTotal + 1;       // 在界内且为故障：计数（In range and faulted, count it）
                            IF nMinPort = 0 THEN
                                nMinPort := p;          // 首次命中即组内最小号（First hit is the lowest port）
                            END_IF
                        END_IF
                    END_IF
                END_FOR
                anGroupMaskOut[g] := uBuildMask;        // 屏蔽后掩码出口（Sanitised mask outlet）
                IF (anGroupFirstPort[g] > 0) AND (anGroupFirstPort[g] <> nMinPort) THEN
                    bPortDeclMismatch := TRUE;          // 声明值与推导值不一致：标记 014C（Declared value differs, flag 014C）
                END_IF
            ELSE
                anGroupMaskOut[g] := DL_MASK_NONE;      // 未启用组掩码清零（Unused group mask cleared）
            END_IF
        END_FOR
        nTotalFaultPort := nTotal;              // 故障总数出口（Fault total outlet）
        bAnyFault       := (nTotal > 0);        // 存在故障（Any fault present）
        (* ② 首出仲裁：仅未锁存时执行，组号优先、端口号次之，取字典序最小 *)
        nGuard := 0;                            // 子段守卫清零（Guard reset for this pass）
        IF (NOT stBoard.bLatchValid) AND (nTotal > 0) THEN
            bFound      := FALSE;               // 命中标志预清零（Hit flag pre-cleared）
            nScanGroup  := 0;                   // 仲裁组号预清零（Arbitration group pre-cleared）
            nScanPort   := 0;                   // 仲裁端口号预清零（Arbitration port pre-cleared）
            FOR g := 1 TO nGroupUse DO
                nGuard := nGuard + 1;           // 守卫递增（Guard incremented）
                IF nGuard > DL_GUARD_MAX THEN
                    EXIT;                       // 守卫到顶即退出（Bail out at the guard bound）
                END_IF
                FOR p := 1 TO auPortCntUse[g] DO
                    nGuard := nGuard + 1;       // 守卫递增（Guard incremented）
                    IF nGuard > DL_GUARD_MAX THEN
                        EXIT;                   // 守卫到顶即退出（Bail out at the guard bound）
                    END_IF
                    IF (NOT bFound) AND ((anGroupMaskOut[g] AND SHL(DL_MASK_ONE, p - 1)) <> DL_MASK_NONE) THEN
                        bFound      := TRUE;    // 命中即锁存（Latch on the first hit）
                        nScanGroup  := g;       // 记录组号（Record the group）
                        nScanPort   := p;       // 记录端口号（Record the port）
                    END_IF
                END_FOR
            END_FOR
            IF bFound THEN
                stBoard.nLatchedGroup := nScanGroup;                  // 锁存组号（Latch the group）
                stBoard.nLatchedPort  := nScanPort;                   // 锁存端口号（Latch the port）
                stBoard.uLatchedCode  := auGroupFirstCode[nScanGroup]; // 组内首出码代表该组（The group first-out code represents the group）
                stBoard.bLatchValid   := TRUE;                        // 置锁存有效（Mark the latch valid）
            END_IF
        END_IF
        (* ③ 待修排序：与仲裁同一字典序，取前三位，空位填 0 *)
        nGuard := 0;                            // 子段守卫清零（Guard reset for this pass）
        nTopCount := 0;                         // 已填位个数清零（Filled slot count cleared）
        FOR g := 1 TO nGroupUse DO
            nGuard := nGuard + 1;               // 守卫递增（Guard incremented）
            IF nGuard > DL_GUARD_MAX THEN
                EXIT;                           // 守卫到顶即退出（Bail out at the guard bound）
            END_IF
            FOR p := 1 TO auPortCntUse[g] DO
                nGuard := nGuard + 1;           // 守卫递增（Guard incremented）
                IF nGuard > DL_GUARD_MAX THEN
                    EXIT;                       // 守卫到顶即退出（Bail out at the guard bound）
                END_IF
                IF (nTopCount < DL_TOP_N) AND ((anGroupMaskOut[g] AND SHL(DL_MASK_ONE, p - 1)) <> DL_MASK_NONE) THEN
                    nTopCount := nTopCount + 1;                        // 占一个待修位（Occupy one slot）
                    anTopPortNo[nTopCount]   := g * DL_GROUP_STRIDE + p; // 编码：组号乘十加端口号（Encode as group times ten plus port）
                    auTopPortCode[nTopCount] := auGroupFirstCode[g];    // 诊断码取组内首出码（Code taken from the group first-out code）
                END_IF
            END_FOR
        END_FOR
        FOR p := 1 TO DL_TOP_N DO
            IF p > nTopCount THEN
                anTopPortNo[p]   := 0;          // 不足三位填空位（Empty slot marked zero）
                auTopPortCode[p] := 0;          // 空位码清零（Empty slot code cleared）
            END_IF
        END_FOR
        (* ④ 掩码跳变风暴：单拍变化位数超阈值只作趋势提示，不锁存、不置故障位 *)
        nGuard := 0;                            // 子段守卫清零（Guard reset for this pass）
        IF bMaskBase THEN
            FOR g := 1 TO DL_GROUP_MAX DO
                uDiff := anGroupMaskOut[g] XOR stBoard.anLastMask[g]; // 掩码差分（Mask difference）
                FOR p := 1 TO DL_PORT_MAX DO
                    IF (uDiff AND SHL(DL_MASK_ONE, p - 1)) <> DL_MASK_NONE THEN
                        nBitScan := nBitScan + 1;   // 变化位计数（Changed bit counted）
                    END_IF
                END_FOR
            END_FOR
            IF nBitScan > DL_JUMP_MAX THEN
                bMaskJump := TRUE;              // 超阈值：标记趋势码 030B（Above the threshold, flag trend code 030B）
            END_IF
        END_IF
        FOR g := 1 TO DL_GROUP_MAX DO
            stBoard.anLastMask[g] := anGroupMaskOut[g]; // 判读完再装载新基准（Load the baseline after the comparison）
        END_FOR
        bMaskBase := TRUE;                      // 基准已就绪（Baseline ready）
        ePhase    := E_DL_BoardPhase.eIdle;     // 本拍结束回待机，无长驻态（Back to idle, never resident）

    E_DL_BoardPhase.eFault: // 故障：输出保持，等复位沿（Fault, outputs held until the reset edge）
        bAnyFault := (nTotalFaultPort > 0);     // 故障位保持期间派生量仍可读（Derived flag stays readable）

    ELSE
        bFaultLatch := TRUE;                    // 非法状态兜底锁存（Illegal state latched）
        uErrInt     := 16#0003_030C;            // 030C 非法状态兜底（Illegal state fallback code）
        ePhase      := E_DL_BoardPhase.eFault;  // 进终端安全态（Enter the terminal safe state）
END_CASE

(*------------------------------------------------------------------------------
 * 段 5｜首出换出（锁存值转出到引脚，复位分支在本段之后执行）
 *      First-out outlet mapping, the reset block runs after this section
 *-----------------------------------------------------------------------------*)
nFirstGroup := stBoard.nLatchedGroup;           // 首出组号出口（First-out group outlet）
nFirstPort  := stBoard.nLatchedPort;            // 首出端口号出口（First-out port outlet）
uFirstCode  := stBoard.uLatchedCode;            // 首出码出口（First-out code outlet）

(*------------------------------------------------------------------------------
 * 段 6｜复位（置于仲裁与换出之后，保证复位当拍首出即为空，下一拍重新仲裁）
 *      Reset runs after arbitration and outlet mapping, so the first-out is empty
 *      on the reset cycle and re-arbitrated on the next one
 *-----------------------------------------------------------------------------*)
IF fbTrigReset.Q THEN
    stBoard.nLatchedGroup := 0;                 // 清锁存组号（Clear the latched group）
    stBoard.nLatchedPort  := 0;                 // 清锁存端口号（Clear the latched port）
    stBoard.uLatchedCode  := 0;                 // 清锁存码（Clear the latched code）
    stBoard.bLatchValid   := FALSE;             // 清锁存有效位（Clear the latch valid flag）
    nFirstGroup           := 0;                 // 复位当拍首出为空（First-out empty on the reset cycle）
    nFirstPort            := 0;                 // 复位当拍首出为空（First-out empty on the reset cycle）
    uFirstCode            := 0;                 // 复位当拍首出码为空（First-out code empty on the reset cycle）
    bFaultLatch           := FALSE;             // 清故障锁存（Clear the fault latch）
    uErrInt               := 16#0000_0000;      // 清故障码（Clear the fault code）
    IF ePhase = E_DL_BoardPhase.eFault THEN
        ePhase := E_DL_BoardPhase.eIdle;        // 故障态复位回待机（Fault returns to idle）
    END_IF
END_IF

(*------------------------------------------------------------------------------
 * 段 7｜码位定级（单一优先级链，全拍只写一次 uErrorId）
 *      Single priority chain, the event code is written once per scan
 *-----------------------------------------------------------------------------*)
IF bMaskJump THEN
    uInfoCode := 16#0003_030B;                  // 优先级一：掩码跳变风暴，仅趋势提示（Mask burst, trend only）
ELSIF bMaskClamped THEN
    uInfoCode := 16#0003_014B;                  // 优先级二：超界位被屏蔽（Out-of-range bits suppressed）
ELSIF bPortDeclMismatch THEN
    uInfoCode := 16#0003_014C;                  // 优先级三：声明首出端口不一致（Declared first-out port mismatch）
ELSIF bGroupClamped THEN
    uInfoCode := 16#0003_0149;                  // 优先级四：组数超上限已钳位（Group count clamped）
ELSIF bPortClamped THEN
    uInfoCode := 16#0003_014A;                  // 优先级五：端口数超上限已钳位（Port count clamped）
ELSIF bGroupShort THEN
    uInfoCode := 16#0003_0309;                  // 优先级六：组数小于 1（Group count below one）
ELSIF bPortShort THEN
    uInfoCode := 16#0003_030A;                  // 优先级七：端口数小于 1（Port count below one）
ELSE
    uInfoCode := 16#0000_0000;                  // 无事件（No event）
END_IF

eState := ePhase;                               // 相位出口（Phase outlet）
bError := bFaultLatch;                          // 故障位只反映故障级锁存（Fault bit reflects the latch only）
IF bFaultLatch THEN
    uErrorId := uErrInt;                        // 故障级码优先透出（Fault level code has priority）
ELSE
    uErrorId := uInfoCode;                      // 无故障透出本拍信息级码（Info code exposed otherwise）
END_IF
END_FUNCTION_BLOCK

(* ---- FB_DL_RefDefrostCycleSeq.st ---- *)
(*
  ============================================================
  组件名 : FB_DL_RefDefrostCycleSeq
  分类   : DL_Device
  功能   : 冷风机除霜循环（制冷 → 判霜 → 融霜 → 滴水 → 恢复），含融霜超时、恢复超时、风机反馈丢失、参数非法四类故障锁存与除霜次数累计
  开源溯源 : internal-design（本轮无外部代码逐行引用）；参考语义 : 无外部参考
  复杂度 : C4
  版本   : 1.0.0
  ============================================================
*)

(*-----------------------------------------------------------------------------
 * 状态迁移表（ENUM 成员 → 出口；每成员均有可到达出口，零无界驻留相）：
 *   eIdle       → eCooling    : bEnable 且组态闸通过且无锁存
 *   eIdle       ── 保持，直到使能（待机相以使能为唯一出口，属许可型驻留）
 *   eCooling    → eFrostDetect: tonCoolMin.Q（已累计满足最短制冷 tCoolMin 才允许判霜）
 *   eCooling    → eIdle       : bEnable 撤除（段 5 失能迁相）
 *   eCooling    → eFault      : tonFanFb.Q（码 3 风机反馈与指令不符）｜组态失效（码 4）
 *   eFrostDetect→ eDefrost    : 判霜判据成立（室温-盘管温差 > 阈值 且 盘管 < 0 且 吸气压力 > 下限）
 *   eFrostDetect→ eCooling    : 判霜判据不成立（本相为单拍决策相，无驻留）
 *   eDefrost    → eDrip       : rCoilTempC ≥ rDefrostTermTempC（达融霜终止温度）
 *   eDefrost    → eFault      : tonDefrost.Q（码 1 融霜超时）｜tonFanFb.Q（码 3）｜bEnable 撤除（段 5）
 *   eDrip       → eRecover    : tonDrip.Q（滴水计时到，本相为定时驻留，出口由计时器保证）
 *   eDrip       → eIdle/eFault: bEnable 撤除（段 5）｜tonFanFb.Q（码 3）
 *   eRecover    → eCooling    : 盘管温度回落至（室温 - 阈值）以下，压缩机延时启动条件成立
 *   eRecover    → eFault      : tonRecover.Q（码 2 恢复超时）｜tonFanFb.Q（码 3）｜bEnable 撤除（段 5）
 *   eFault      → eIdle       : bEnable 重新使能的上升沿（下降沿后再使能，段 3 分支内清锁存）
 *   ELSE（非法枚举值，非任何成员）→ eFault（码 5）
 *
 * 故障码表（nFaultCode，0 = 无故障；非首码均附「现有输出不可观测」反证句，R90）：
 *   1 融霜超时   : tonDefrost 覆盖 eDefrost 全相，达 tDefrostMax 仍未到终止温度即锁存。
 *   2 恢复超时   : 反证——恢复相 bCompressorOn = FALSE 而 bFanOn = TRUE，与码 1 的
 *                  「风机与压缩机全关」时序签名不同；但故障相动作全撤后两者观测量一致，
 *                  复用码 1 会把「融霜水未排干/盘管未回落」误报为「加热不足」，处置方向相反。
 *   3 风机反馈失 : 反证——反馈丢失可由 eCooling（应转却在停）与 eDefrost（应停却在转）两侧触发，
 *                  与任何超时码无共享观测量；复用超时码会让机械故障被当作时间参数问题。
 *   4 参数非法   : 反证——非法阈值/时间在启动瞬间拦截，无除霜动作、无计数递增，
 *                  与码 1/2/3 的时序签名互斥，必须独立成码以便组态错误可前置观测。
 *   5 非法状态   : 反证——非法枚举值为程序缺陷而非现场事件，合并入任一工艺码会让
 *                  固件错误被误排为制冷系统故障，必须独立成码。
 *
 * 依赖     : 仅 IEC 61131-3 标准库（TON / R_TRIG / ABS），零厂商私有库
 * 分工声明 : 压缩机高低压保护与吸气压力联锁归压缩机组保护件；本件只做除霜时序、
 *            风机反馈一致性监视与除霜次数累计，不做制冷量调节、不做电机过载保护。
 *            吸气压力在本件只作判霜前置闸（系统未运行时禁止判霜），不作保护判据。
 * 归属     : E_DL_RefDfsState 归属本文件（全库唯一定义，R264；引用件只引用不重声明）。
 * 修订历史 : 2026-11-25  v1.0.0  首版（编码席 dlf-plc-coder，第二批 C4）
 *----------------------------------------------------------------------------*)

(*-----------------------------------------------------------------------------
 * 边界与红线自检：
 * ① 五个 TON 与一个 R_TRIG 全部在 CASE 外无条件周期调用（R7）；时间类 IN 均含 NOT .Q 自复位项
 *    与 NOT 故障锁存项（R188 / FB50-1③），CASE 内只读 .Q。
 * ② 三个执行出口（压缩机 / 除霜阀 / 风机）在段 0 每拍预置 FALSE，CASE 内只置 TRUE；
 *    段 5 在 eIdle 与 eFault 相再次全撤 —— eIdle 三输出必为 FALSE，无上一相残留。
 * ③ 风机反馈判据用「相位期望值」比较（R99 状态量门控），不用上一拍命令位：期望为真的相
 *    为 eCooling / eFrostDetect / eRecover，期望为假的相为 eIdle / eDefrost / eDrip / eFault；
 *    不符持续 DL_DFS_FB_WIN（3s）才置码 3，避开启动/停止瞬间的机械过渡。
 * ④ 除霜次数 _nCount 只在 eFrostDetect → eDefrost 迁移点 +1（单点写入，一霜一次）；
 *    本件任何复位路径都不清零该计数（FB50-2② 作用域声明：由上层维护清零）。
 * ⑤ 复位沿作用域（FB50-2②）：eFault 内 bEnable 上升沿 = 清故障锁存 + 清故障码 + 迁相回 eIdle，
 *    三项各写明；bEnable 下降沿的作用域 = 迁相回 eIdle 并全撤输出，不清锁存、不清计数。
 * ⑥ 组态域闸枚举全部浮点入参（rCoilTempC / rRoomTempC / rSuctionPressBar / rFrostThresh /
 *    rDefrostTermTempC），NaN 自反 + Inf 差值自减双判（R151 / R79）。
 * ⑦ 零全局耦合：无 GVL / VAR_EXTERNAL / %I / %Q（R1 / R2）；无 FOR / WHILE / REPEAT（R271 N/A）。
 * ⑧ 相位写入点共两处且互斥：段 3 CASE、段 5 段尾迁移闸。
 *----------------------------------------------------------------------------*)

TYPE E_DL_RefDfsState :
(
    eIdle        := 0,                                              // 空闲：压缩机/除霜阀/风机全停，等使能 idle: compressor, defrost valve and fan all off, waiting for enable
    eCooling     := 1,                                              // 制冷相：压缩机与风机开，累计最短制冷时间 cooling: compressor and fan on, accumulating the minimum cooling time
    eFrostDetect := 2,                                              // 判霜决策相：单拍决策，不改变执行出口 frost detect: single scan decision without changing the actuators
    eDefrost     := 3,                                              // 融霜相：压缩机关、除霜阀开、风机关，至终止温度 defrost: compressor off, defrost valve on, fan off until the termination temperature
    eDrip        := 4,                                              // 滴水相：三输出全关，等 tDripTime drip: all three outputs off until tDripTime elapses
    eRecover     := 5,                                              // 恢复相：风机先开，盘管回落后压缩机延时启动 recover: fan first, the compressor starts after the coil recovers
    eFault       := 6                                               // 故障锁存相：三输出全停，只由 bEnable 重新使能迁出 fault: all outputs off, left only by a re-enabled bEnable
);
END_TYPE

FUNCTION_BLOCK FB_DL_RefDefrostCycleSeq
VAR_INPUT
    bEnable           : BOOL := FALSE;                              // 除霜循环使能（电平）：撤除即三输出全停 [bool] defrost cycle enable level, dropping it stops all outputs
    rCoilTempC        : REAL := 0.0;                                // 盘管表面实测温度 [degC] measured coil surface temperature [degC]
    rRoomTempC        : REAL := 0.0;                                // 库房空气实测温度 [degC] measured room air temperature [degC]
    rSuctionPressBar  : REAL := 0.0;                                // 压缩机吸气压力 [bar] compressor suction pressure [bar]
    bFanFeedback      : BOOL := FALSE;                              // 风机运行反馈（TRUE = 在转）[bool] fan running feedback, TRUE means running
    rFrostThresh      : REAL := 5.0;                                // 判霜温差阈值（室温-盘管），域 > 0 [K] frost detection temperature difference threshold, domain > 0 [K]
    rDefrostTermTempC : REAL := 8.0;                                // 融霜终止温度（盘管回升到此值即结束），域 > 0 [degC] defrost termination coil temperature, domain > 0 [degC]
    tDefrostMax       : TIME := T#20M;                              // 融霜最长时长 [s] maximum defrost duration [s]
    tDripTime         : TIME := T#3M;                               // 滴水时长（融霜后滴排残水）[s] drip duration after defrost [s]
    tRecoverMax       : TIME := T#10M;                              // 恢复最长时长 [s] maximum recovery duration [s]
    tCoolMin          : TIME := T#15M;                              // 最短制冷时长（满足后才允许判霜）[s] minimum cooling time before frost detection is allowed [s]
END_VAR
VAR_OUTPUT
    bCompressorOn    : BOOL;                                        // 压缩机运行命令（段 0 预置，CASE 只置位）[bool] compressor run command
    bDefrostValveOn  : BOOL;                                        // 除霜阀命令（仅融霜相）[bool] defrost valve command, defrost phase only
    bFanOn           : BOOL;                                        // 风机运行命令（制冷/判霜/恢复相）[bool] fan run command in cooling, detect and recovery phases
    eState           : E_DL_RefDfsState;                            // 相位出口（段 6 单点映射）[-] phase outlet mapped once in section 6
    nDefrostCount    : INT;                                         // 累计除霜次数（本件不清零，由上层维护）[次] accumulated defrost count maintained by the upper layer
    bDefrostAlarm    : BOOL;                                        // 除霜告警（故障锁存派生位，需人工/复位确认）[bool] defrost alarm derived from the fault latch
    nFaultCode       : INT;                                         // 故障码 0 无 1 融霜超时 2 恢复超时 3 风机反馈丢失 4 参数非法 5 非法状态 [码] fault code
    bError           : BOOL;                                        // 故障锁存标志（取锁存位，R45 配对出口）[bool] fault latch flag used as the paired outlet
END_VAR
VAR
    _eState      : E_DL_RefDfsState := E_DL_RefDfsState.eIdle;      // 内部相位（CASE 唯一比较目标）[-] internal phase compared by the CASE
    _bFaultLatch : BOOL := FALSE;                                   // 故障锁存位（仅 bEnable 重新使能沿清除）[bool] fault latch, cleared only by a re-enabled bEnable edge
    _nFault      : INT := 0;                                        // 锁存故障码（故障期回放，不按当下输入重算）[码] latched fault code replayed in the fault phase
    _nCount      : INT := 0;                                        // 内部除霜次数累计（单点写入）[次] internal defrost count with a single write point
    _bCfgOk      : BOOL := FALSE;                                   // 组态与入参域闸通过标志 [bool] configuration and input domain gate flag
    _bRunActive  : BOOL := FALSE;                                   // 制冷相关相标志（制冷到恢复）[bool] cooling related phase flag from cooling to recovery
    _bComp       : BOOL := FALSE;                                   // 内部压缩机命令状态 [bool] internal compressor command state
    _bDfv        : BOOL := FALSE;                                   // 内部除霜阀命令状态 [bool] internal defrost valve command state
    _bFan        : BOOL := FALSE;                                   // 内部风机命令状态 [bool] internal fan command state
    _bFanExpect  : BOOL := FALSE;                                   // 按相位推导的风机应有状态（R99 状态量门控）[bool] fan state expected from the phase
    _bFanMismatch : BOOL := FALSE;                                  // 风机反馈与期望不符标志 [bool] fan feedback mismatching the expectation
    rtEnable     : R_TRIG;                                          // bEnable 上升沿实例（段 2 无条件调用）[bool] enable rising edge instance
    tonCoolMin   : TON;                                             // 最短制冷计时（段 2 无条件调用）[s] minimum cooling timer
    tonDefrost   : TON;                                             // 融霜最长时长计时（段 2 无条件调用）[s] maximum defrost timer
    tonDrip      : TON;                                             // 滴水时长计时（段 2 无条件调用）[s] drip timer
    tonRecover   : TON;                                             // 恢复最长时长计时（段 2 无条件调用）[s] maximum recovery timer
    tonFanFb     : TON;                                             // 风机反馈不符持续计时（段 2 无条件调用）[s] fan feedback mismatch persistence timer
END_VAR
VAR CONSTANT
    DL_DFS_ZERO      : REAL := 0.0;                                 // 浮点零基准（亦作盘管结霜温度界限）[degC] float zero base, also the coil frosting limit [degC]
    DL_DFS_PRESS_MIN : REAL := 0.1;                                 // 吸气压力下限（系统运行判据）[bar] suction pressure lower bound proving the system runs [bar]
    DL_DFS_FB_WIN    : TIME := T#3S;                                // 风机反馈不符持续判窗 [s] fan feedback mismatch persistence window [s]
    DL_DFS_T_MIN     : TIME := T#100MS;                             // 时间参数下限 [s] lower bound of the time parameters
    DL_DFS_T_MAX     : TIME := T#8H;                                // 时间参数上限 [s] upper bound of the time parameters
    DL_DFS_CNT_ONE   : INT := 1;                                    // 计数步长 [次] count step
END_VAR

(* —— 段 0：出口预置与派生量（CASE 内只置 TRUE，eIdle / eFault 零残留） —— *)
_bComp := FALSE;                                                    // 压缩机命令每拍先撤 [bool] compressor command withdrawn first each scan
_bDfv  := FALSE;                                                    // 除霜阀命令每拍先撤 [bool] defrost valve command withdrawn first each scan
_bFan  := FALSE;                                                    // 风机命令每拍先撤 [bool] fan command withdrawn first each scan
_bRunActive := (_eState = E_DL_RefDfsState.eCooling) OR (_eState = E_DL_RefDfsState.eFrostDetect)
               OR (_eState = E_DL_RefDfsState.eDefrost) OR (_eState = E_DL_RefDfsState.eDrip)
               OR (_eState = E_DL_RefDfsState.eRecover);            // 制冷相关相标志（用状态量，R99）[bool] cooling related phase flag
_bFanExpect := (_eState = E_DL_RefDfsState.eCooling) OR (_eState = E_DL_RefDfsState.eFrostDetect)
               OR (_eState = E_DL_RefDfsState.eRecover);            // 风机应有状态（按相位推导）[bool] fan state expected from the phase
_bFanMismatch := _bRunActive AND _bFanExpect AND (NOT bFanFeedback); // 反馈不符（只监视「应转未转」，见 R80 闸 B MAJOR-1）[bool] mismatch only when fan expected on

(* —— 段 1：组态域闸（五个浮点入参全枚举，非有限双判 R151 / R79） —— *)
_bCfgOk := TRUE;                                                    // 组态闸标志初值 [bool] configuration flag initial value
IF (rCoilTempC <> rCoilTempC) OR ((rCoilTempC - rCoilTempC) <> DL_DFS_ZERO)
   OR (rRoomTempC <> rRoomTempC) OR ((rRoomTempC - rRoomTempC) <> DL_DFS_ZERO)
   OR (rSuctionPressBar <> rSuctionPressBar) OR ((rSuctionPressBar - rSuctionPressBar) <> DL_DFS_ZERO)
   OR (rFrostThresh <> rFrostThresh) OR ((rFrostThresh - rFrostThresh) <> DL_DFS_ZERO)
   OR (rDefrostTermTempC <> rDefrostTermTempC) OR ((rDefrostTermTempC - rDefrostTermTempC) <> DL_DFS_ZERO) THEN
    _bCfgOk := FALSE;                                               // 非有限入参：拒收（NaN 自反 + Inf 差值自减）[bool] non finite input rejected
END_IF
IF _bCfgOk THEN
    IF rFrostThresh <= DL_DFS_ZERO THEN
        _bCfgOk := FALSE;                                           // 判霜阈值非正（永不判霜）[bool] non positive frost threshold
    ELSIF rDefrostTermTempC <= DL_DFS_ZERO THEN
        _bCfgOk := FALSE;                                           // 终止温度非正（融霜不足）[bool] non positive termination temperature
    ELSIF (tDefrostMax < DL_DFS_T_MIN) OR (tDefrostMax > DL_DFS_T_MAX) THEN
        _bCfgOk := FALSE;                                           // 融霜最长时长越域 [bool] defrost maximum out of domain
    ELSIF (tDripTime < DL_DFS_T_MIN) OR (tDripTime > DL_DFS_T_MAX) THEN
        _bCfgOk := FALSE;                                           // 滴水时长越域 [bool] drip time out of domain
    ELSIF (tRecoverMax < DL_DFS_T_MIN) OR (tRecoverMax > DL_DFS_T_MAX) THEN
        _bCfgOk := FALSE;                                           // 恢复最长时长越域 [bool] recovery maximum out of domain
    ELSIF (tCoolMin < DL_DFS_T_MIN) OR (tCoolMin > DL_DFS_T_MAX) THEN
        _bCfgOk := FALSE;                                           // 最短制冷时长越域 [bool] minimum cooling time out of domain
    END_IF
END_IF
IF (NOT _bCfgOk) AND (NOT _bFaultLatch) AND (bEnable OR _bRunActive) THEN
    _nFault      := 4;                                              // 故障级：参数非法 [码] fault: illegal parameter
    _bFaultLatch := TRUE;                                           // 置故障锁存 [bool] latch the fault
    bError       := TRUE;                                           // R45 配对：故障标志同拍置位 [bool] paired error flag
END_IF

(* —— 段 2：沿与定时器（CASE 外无条件周期调用，R7；IN 含 NOT .Q 自复位与 NOT 锁存，R188） —— *)
rtEnable(CLK := bEnable);                                           // 使能沿无条件刷新 [bool] enable edge refreshed unconditionally
tonCoolMin(IN := (_eState = E_DL_RefDfsState.eCooling) AND (NOT tonCoolMin.Q) AND (NOT _bFaultLatch),
           PT := tCoolMin);                                         // 最短制冷计时 [s] minimum cooling timer
tonDefrost(IN := (_eState = E_DL_RefDfsState.eDefrost) AND (NOT tonDefrost.Q) AND (NOT _bFaultLatch),
           PT := tDefrostMax);                                      // 融霜最长时长 [s] maximum defrost timer
tonDrip(IN := (_eState = E_DL_RefDfsState.eDrip) AND (NOT tonDrip.Q) AND (NOT _bFaultLatch),
        PT := tDripTime);                                           // 滴水时长 [s] drip timer
tonRecover(IN := (_eState = E_DL_RefDfsState.eRecover) AND (NOT tonRecover.Q) AND (NOT _bFaultLatch),
           PT := tRecoverMax);                                      // 恢复最长时长 [s] maximum recovery timer
tonFanFb(IN := _bFanMismatch AND (NOT tonFanFb.Q) AND (NOT _bFaultLatch),
         PT := DL_DFS_FB_WIN);                                      // 风机反馈不符持续判 [s] fan feedback mismatch persistence

(* —— 段 3：主状态机（相位写入点之一；每成员独立标签，ELSE 只兜非法值，FB32-5） —— *)
CASE _eState OF
E_DL_RefDfsState.eIdle :                                            // 空闲相：三输出已撤
    IF bEnable AND _bCfgOk AND (NOT _bFaultLatch) THEN
        _eState := E_DL_RefDfsState.eCooling;                       // 迁移：进入制冷相 [phase] move to cooling
    END_IF

E_DL_RefDfsState.eCooling :                                         // 制冷相：压缩机与风机开
    _bComp := TRUE;                                                 // 压缩机运行 [bool] compressor running
    _bFan  := TRUE;                                                 // 风机运行 [bool] fan running
    IF tonCoolMin.Q THEN
        _eState := E_DL_RefDfsState.eFrostDetect;                   // 迁移：最短制冷已满足，允许判霜 [phase] minimum cooling satisfied, frost detection allowed
    END_IF

E_DL_RefDfsState.eFrostDetect :                                     // 判霜决策相（单拍过渡态）
    (* 拍 N 进入（tonCoolMin.Q 置位）/ 本拍行为：只做判霜决策，执行出口沿用制冷相的安全状态
       （压缩机与风机保持开），不产生任何新动作 / 拍 N+1 转出至 eDefrost 或回 eCooling *)
    _bComp := TRUE;                                                 // 判霜拍沿用压缩机运行 [bool] compressor kept running in the detect scan
    _bFan  := TRUE;                                                 // 判霜拍沿用风机运行 [bool] fan kept running in the detect scan
    IF ((rRoomTempC - rCoilTempC) > rFrostThresh) AND (rCoilTempC < DL_DFS_ZERO)
       AND (rSuctionPressBar > DL_DFS_PRESS_MIN) THEN
        _nCount := _nCount + DL_DFS_CNT_ONE;                        // 除霜次数 +1（单点写入，一霜一次）[次] one count per confirmed frost
        _eState := E_DL_RefDfsState.eDefrost;                       // 迁移：判霜成立进入融霜 [phase] frost confirmed, start the defrost
    ELSE
        _eState := E_DL_RefDfsState.eCooling;                       // 迁移：未达判霜条件回制冷继续累计 [phase] no frost, resume cooling
    END_IF

E_DL_RefDfsState.eDefrost :                                         // 融霜相：压缩机关、除霜阀开、风机关
    _bDfv := TRUE;                                                  // 除霜阀开（压缩机与风机保持关）[bool] defrost valve open
    IF rCoilTempC >= rDefrostTermTempC THEN
        _eState := E_DL_RefDfsState.eDrip;                          // 迁移（出口 1）：盘管达融霜终止温度 [phase] coil reached the termination temperature
    END_IF

E_DL_RefDfsState.eDrip :                                            // 滴水相：三输出全关，等 tDripTime
    IF tonDrip.Q THEN
        _eState := E_DL_RefDfsState.eRecover;                       // 迁移（出口 1）：滴水时间到 [phase] drip time elapsed
    END_IF

E_DL_RefDfsState.eRecover :                                         // 恢复相：风机先开，压缩机延时启动
    _bFan := TRUE;                                                  // 风机先开（化霜水汽排空）[bool] fan first to clear the moisture
    IF rCoilTempC <= (rRoomTempC - rFrostThresh) THEN
        _bComp := TRUE;                                             // 压缩机启动条件成立（盘管已回落）[bool] compressor start condition satisfied
        _eState := E_DL_RefDfsState.eCooling;                       // 迁移（出口 1）：恢复正常制冷 [phase] back to normal cooling
    END_IF

E_DL_RefDfsState.eFault :                                           // 故障锁存相：三输出已由段 5 全撤
    IF rtEnable.Q THEN
        _bFaultLatch := FALSE;                                      // 复位作用域①：清故障锁存（bEnable 下降后再使能的上升沿）[bool] reset scope one
        _nFault      := 0;                                          // 复位作用域②：清故障码 [码] reset scope two
        _eState      := E_DL_RefDfsState.eIdle;                     // 复位作用域③：迁相回空闲 [phase] reset scope three
    END_IF

ELSE                                                                // 非法枚举值兜底（R6 / FB32-5）
    IF NOT _bFaultLatch THEN
        _nFault      := 5;                                          // 故障级：非法状态枚举值 [码] fault: illegal state enum value
        _bFaultLatch := TRUE;                                       // 置故障锁存 [bool] latch the fault
        bError       := TRUE;                                       // R45 配对：故障标志同拍置位 [bool] paired error flag
    END_IF
    _eState := E_DL_RefDfsState.eFault;                             // 非法值一律落安全相 [phase] illegal value falls into the safe phase
END_CASE

(* —— 段 4：超时看门狗锁存（状态已迁出则该相看门狗不生效，R275） —— *)
IF tonDefrost.Q AND (NOT _bFaultLatch) AND (_eState = E_DL_RefDfsState.eDefrost) THEN
    _nFault      := 1;                                              // 故障级：融霜超时未达终止温度 [码] fault: defrost timeout before the termination temperature
    _bFaultLatch := TRUE;                                           // 置故障锁存 [bool] latch the fault
    bError       := TRUE;                                           // R45 配对：故障标志同拍置位 [bool] paired error flag
END_IF
IF tonRecover.Q AND (NOT _bFaultLatch) AND (_eState = E_DL_RefDfsState.eRecover) THEN
    _nFault      := 2;                                              // 故障级：恢复超时 [码] fault: recovery timeout
    _bFaultLatch := TRUE;                                           // 置故障锁存 [bool] latch the fault
    bError       := TRUE;                                           // R45 配对：故障标志同拍置位 [bool] paired error flag
END_IF
IF tonFanFb.Q AND (NOT _bFaultLatch) AND _bRunActive THEN
    _nFault      := 3;                                              // 故障级：风机反馈丢失（与相位期望不符持续 3s）[码] fault: fan feedback lost
    _bFaultLatch := TRUE;                                           // 置故障锁存 [bool] latch the fault
    bError       := TRUE;                                           // R45 配对：故障标志同拍置位 [bool] paired error flag
END_IF

(* —— 段 5：失能迁相 + 段尾故障迁移闸 + 空闲/故障相输出全撤（FB50-1④ / R191 显式声明） —— *)
IF (NOT bEnable) AND (_eState <> E_DL_RefDfsState.eFault) THEN
    (* 失能语义（R191 二选一，本件选「降级为安全值 + 回空闲，不置故障码」）：
       作用域仅迁相位与撤输出，不清故障锁存、不清除霜计数 *)
    _eState := E_DL_RefDfsState.eIdle;                              // 失能即安全停机回空闲 [phase] disable stops safely into idle
END_IF
IF _bFaultLatch AND (_eState <> E_DL_RefDfsState.eFault) THEN
    _eState := E_DL_RefDfsState.eFault;                             // 锁存即迁相（锁存与迁相分离，R21）[phase] a latch forces the fault phase
END_IF
IF (_eState = E_DL_RefDfsState.eIdle) OR (_eState = E_DL_RefDfsState.eFault) THEN
    _bComp := FALSE;                                                // 空闲/故障：压缩机全停 [bool] compressor off in idle and fault
    _bDfv  := FALSE;                                                // 空闲/故障：除霜阀全关 [bool] defrost valve closed in idle and fault
    _bFan  := FALSE;                                                // 空闲/故障：风机全停 [bool] fan off in idle and fault
END_IF

(* —— 段 6：统一出口（执行映射 + 计数 + 告警派生 + 锁存码回放；单点写入） —— *)
bCompressorOn   := _bComp;                                          // 压缩机命令出口 [bool] compressor command outlet
bDefrostValveOn := _bDfv;                                           // 除霜阀命令出口 [bool] defrost valve command outlet
bFanOn          := _bFan;                                           // 风机命令出口 [bool] fan command outlet
eState          := _eState;                                         // 相位出口 [phase] phase outlet
nDefrostCount   := _nCount;                                         // 除霜次数出口 [次] defrost count outlet
bDefrostAlarm   := _bFaultLatch;                                    // 除霜告警取故障锁存位（派生位，R28 5.9）[bool] alarm derived from the fault latch
nFaultCode      := _nFault;                                         // 故障码出口（锁存回放）[码] fault code outlet replayed from the latch
bError          := _bFaultLatch;                                    // 故障标志取锁存位 [bool] fault flag from the latch
END_FUNCTION_BLOCK

(* ---- FB_DL_RollerGapAdjust.st ---- *)
(*==============================================================================
 * 组件名称 (Component)  : FB_DL_RollerGapAdjust
 * 所属子库 (Sublibrary) : DL_Device
 * 当前版本 (Version)    : 1.0.0
 * 组件分类 (Category)   : 功能块（FUNCTION_BLOCK）· 设备执行 · 辊距微调背隙补偿
 * 兼容性   (Platform)   : CODESYS 3.5 / TwinCAT 3 / 汇川 InoProShop / Schneider
 *                         Machine Expert；仅 LIMIT / ABS 与标准 TON / R_TRIG
 * 功能描述 (Function)   : 把「目标辊距 → 单向越程逼近（吃掉背隙）→ 反向精定位
 *                         → 到位窗口判定 → 偏差记账」封装成设备对象，输出电动
 *                         缸位置指令与到位状态。解决电动缸双向逼近时背隙导致
 *                         的重复定位偏差，让每次调整都从同一侧逼近目标。
 * 边界声明 (Boundary)   : FB_DL_ThreePointValve 是浮点式阀的开度积分估算；
 *                         FB_DL_AnalogValve 是模拟量比例阀开度控制；本块是
 *                         位置伺服式间隙调整（带背隙补偿与到位窗口）。三者执行
 *                         机构语义不同，不可互替。本块刻意不注入轴接口：辊距
 *                         调整多为独立电动缸加位移传感器，注入轴接口会把设备层
 *                         拖到运动层，破坏分层依赖方向。
 * 为什么必须两段     : 单向逼近是背隙补偿的本体。把两段压成「一次赋值加到位
 *                     判定」会丢掉「先越程再回退」的动作序列，重复定位精度退化
 *                     到双向逼近水平——那正是普通定位块已有的能力，本件也就没有
 *                     存在价值。故 eApproach 与 eFine 是不可合并的两个相位。
 * 背隙补偿算术   : 阶段 A 指令取「目标加逼近符号乘背隙」，逼近符号为负一，
 *                     即先退到目标下方一个背隙；反馈越程过半后进入阶段 B，
 *                     指令回目标值，反向逼近吃掉整段背隙。两个阶段都必须把
 *                     指令钳在上下限内，防止背隙量把指令推出机械行程。
 * 反馈丢失纪律   : 位移反馈无效时指令必须**保持上一拍值**，绝不清零——对辊距
 *                     来说指令清零等于辊缝全开，属于危险侧动作。同时撤回到位
 *                     标志（位置不可信），并置反馈丢失故障码，等待人工确认。
 * 到位与记账     : 到位判定同时要求「偏差在容差内」与「反馈有效」，两者缺一
 *                     不可；到位拍写残余偏差、更新偏差一阶低通均值、更新本次
 *                     调整耗时，并对超容差次数累加。统计量用于预测机械磨损。
 * 开源溯源 (Origin)   : rockwell-aoi / lbp-process / lgf-technology。参考公开
 *                     设备 AOI 的参数分段组织与工艺功能库中「单向逼近消除背隙」
 *                     的工艺分类，只借参数分段与工艺分类；状态机、指令算术、
 *                     钳位策略、统计口径、码位与全部实现 100% 自有，clean-room
 *                     实现，不构成衍生作品。
 * 依赖     (Depends)   : 无 DL_ 内部依赖；仅 Standard.library 的 TON / R_TRIG
 * 故障码表 (Error codes):
 *   16#0003_0147【信息级】目标间隙越界已钳位（含上下限颠倒时的自动换位）
 *   16#0003_0148【信息级】背隙补偿量越界已钳位（负值或超上限）
 *   16#0003_0305【故障级】到位超时（限时内偏差始终未进入容差带）
 *   16#0003_0306【故障级】位移反馈无效或丢失（指令保持，撤回到位标志）
 *   16#0003_0308【故障级】非法相位兜底
 * 码位占用 (Slot)      : 信息级 0147 / 0148；故障级 0305 / 0306 / 0308。
 *                         全部落在 R11 本件分配块内，无跨块借用。
 * 写入点次序 (Write order) :
 *   ① fGapCmd    ：只在相位跃迁拍写（进逼近写越程值，进精定位写目标值），
 *                  其余拍一律不写，从而天然满足「故障时指令保持」
 *   ② bInPosition：只在到位跃迁拍置真，启动新一次调整时置假，其余拍不写
 *   ③ ePhase     ：状态机段为唯一位移点，复位分支只回待机
 *   ④ uErrorId   ：输出段单一优先级链（0308 优于 0306 优于 0305 优于 0147
 *                  优于 0148），全拍只写一次
 * 验收向量 (Acceptance) :
 *   V1 两阶段指令：目标 2.500、背隙 0.050 → 阶段 A 指令 2.450；到位保持段 2.500
 *   V2 到位判定：目标 2.500、容差 0.02、反馈 2.515 → 到位为真、残余偏差 +0.015
 *   V3 限幅：目标 5.0、上限 3.0 → 钳位后阶段 A 指令落在 2.950，保持段指令 3.000，
 *      并置码 16#0003_0147
 *   V4 反馈丢失：反馈有效由真变假（指令原为 2.50）→ 指令保持 2.50、码
 *      16#0003_0306、故障位为真
 *   V5 超时：限时 10 秒内偏差始终大于容差 → 码 16#0003_0305、调整中为假、
 *      累计调整次数不加
 * 红线自检 (Redline)   : R1 零全局变量表与外部变量引用 ｜ R2 零物理地址直写
 *                        R3 纯 IEC 61131-3 ｜ R4 浮点全用容差比较、无除法
 *                        R5 全变量中英双语同行注释 ｜ R6 ENUM 加 CASE 加 ELSE
 *                        R7 TON 与两个 R_TRIG 在 CASE 之外无条件刷新
 *                        R8 信息级码 0147 与 0148 不置故障位
 * 修订历史 (Revision)  :
 *   2026-11-15  v1.0.0  首版落盘（Round 11 · 泳道 B · 辊距伺服微调）
 *============================================================================*)

(*------------------------------------------------------------------------------
 * 结构体: ST_DL_GapTrimStat（跨周期统计，由调用方持有）
 *         Persistent statistics structure owned by the caller
 *-----------------------------------------------------------------------------*)
TYPE ST_DL_GapTrimStat :
STRUCT
    fDevAvg    : REAL;      // 残余偏差一阶低通均值 [毫米]，用于预测机械磨损 / Low pass average of the residual deviation, millimetre
    tLastMove  : TIME;      // 上一次调整的耗时 [毫秒] / Duration of the last adjustment
    nOverTolCnt : UDINT;    // 偏差超容差次数，饱和计数 [次] / Count of adjustments that ended outside the tolerance band
END_STRUCT
END_TYPE

(*------------------------------------------------------------------------------
 * 枚举: E_DL_GapPhase（本块相位，归属本功能块并同文件发布）
 *       Phase enumeration owned by this block and published in the same file
 *-----------------------------------------------------------------------------*)
TYPE E_DL_GapPhase :
(
    eIdle     := 0,   // 待机：可接受启动沿，指令保持 / Idle, ready for a start edge, command kept
    eApproach := 10,  // 逼近：先越程一个背隙，从同一侧靠近 / Approach, overshoot by one backlash from one side
    eFine     := 20,  // 精定位：反向逼近到目标值 / Fine positioning, approach the target from the opposite side
    eHold     := 30,  // 保持：到位后维持指令，等待下一次调整 / Hold, keep the command until the next adjustment
    eFault    := 99   // 故障：超时或反馈丢失，需复位 / Fault, timeout or feedback loss, needs a reset
);
END_TYPE

(*==============================================================================
 * 逐拍推演 (Cycle-by-cycle trace)：
 *   场景 A 正常一次调整（目标 2.500，背隙 0.050，容差 0.02）
 *     启动沿拍：反馈有效，进逼近相位，指令写 2.450，到位标志清假，限时开始计时
 *     逼近相位：段五算出越程过半判据点为 2.475，反馈降到 2.470 时进精定位，
 *          指令改写 2.500
 *     精定位相位：反馈升到 2.515，偏差 0.015 在容差内，进保持相位，到位置真，
 *          残余偏差写 0.015，偏差均值按低通系数更新，耗时取限时器已计时间
 *     保持相位：指令维持 2.500，不再改写；下一次启动沿才重新走两段
 *   场景 B 到位超时（限时十秒，偏差始终 0.5 毫米）
 *     精定位相位中限时器到拍：转故障相位，码 0305，调整中标志落，累计调整
 *     次数不加（未到位不计入台账）
 *   场景 C 反馈丢失（指令原为 2.500）
 *     反馈有效位变假：逼近与精定位相位转故障，保持相位只报警不断开保持；
 *     指令**不写**，自然保持 2.500；到位标志撤回；码 0306
 *   场景 D 目标越界（目标 5.0，上限 3.0）
 *     段三先钳位目标到 3.0 并标记，段四的上下限颠倒检查确认顺序正确；
 *     指令装配时再钳一次，保证背隙量不会把指令推出机械行程；码 0147 只进码
 *   场景 E 非法相位（枚举被外部强制写成未定义值）
 *     兜底分支转故障相位并置 0308，指令保持，需复位退出
 *============================================================================*)

FUNCTION_BLOCK FB_DL_RollerGapAdjust
VAR_INPUT
    bEnable        : BOOL;                  // 使能，FALSE 时指令保持、撤回到位标志 [-] / Enable, holds the command and drops the in-position flag
    bReset         : BOOL;                  // 复位故障，上升沿有效 [-] / Clears the fault on a rising edge
    bAdjustStart   : BOOL;                  // 执行一次调整，上升沿触发 [-] / Triggers one adjustment on a rising edge
    fGapSetpoint   : REAL;                  // 目标辊距 [毫米]，量程 0.0 到 20.0 / Target roller gap in millimetre, zero to twenty
    fGapActual     : REAL;                  // 位移传感器实测辊距 [毫米] / Measured roller gap in millimetre
    fGapTol        : REAL := 0.02;          // 到位容差 [毫米]，0 表示必须完全相等 / In-position tolerance in millimetre, zero demands equality
    fBacklash      : REAL := 0.05;          // 反向背隙补偿量 [毫米]，0 表示不补偿 / Backlash compensation in millimetre, zero disables it
    fCmdMin        : REAL := 0.0;           // 指令下限 [毫米] / Command lower limit in millimetre
    fCmdMax        : REAL := 20.0;          // 指令上限 [毫米] / Command upper limit in millimetre
    bFeedbackValid : BOOL;                  // 位移反馈有效（传感器自诊断汇总）[-] / Position feedback valid, sensor self diagnosis summary
    tMoveTimeout   : TIME := T#10S;         // 单次调整限时 [毫秒]，0 表示不监控 / Adjustment timeout, zero disables monitoring
END_VAR
VAR_OUTPUT
    fGapCmd        : REAL;                  // 电动缸位置指令 [毫米]，故障时保持不写 / Actuator position command, kept untouched on a fault
    bAdjusting     : BOOL;                  // 调整进行中（逼近或精定位）[-] / Adjustment in progress, approach or fine
    bInPosition    : BOOL;                  // 到位，保持到下次调整 [-] / In position, kept until the next adjustment
    eState         : E_DL_GapPhase;         // 主状态机当前相位 [-] / Current phase of the main state machine
    bError         : BOOL;                  // 故障级锁存，仅 0305 0306 0308 置位 [-] / Latched fault, only fault level codes set it
    uErrorId       : UDINT;                 // 事件码，0 表示无事件 [代码] / Event code, zero means none
    fLastDeviation : REAL;                  // 上次调整结束时的残余偏差 [毫米] / Residual deviation of the last adjustment
    nAdjustCount   : UDINT;                 // 累计调整次数，仅到位时累加，饱和 [次] / Adjustment counter, saturating, incremented on arrival only
END_VAR
VAR_IN_OUT
    stTrim         : ST_DL_GapTrimStat;     // 跨周期统计：偏差均值、耗时、超容差次数 / Persistent statistics, deviation, duration and over tolerance count
END_VAR
VAR
    fbTrigReset    : R_TRIG;                // 复位沿检测，CASE 之外无条件刷新 [-] / Reset edge detector, refreshed outside the CASE
    fbTrigStart    : R_TRIG;                // 启动沿检测，CASE 之外无条件刷新 [-] / Start edge detector, refreshed outside the CASE
    fbTonMove      : TON;                   // 单次调整限时计时，CASE 之外无条件刷新 / Move timeout timer, refreshed outside the CASE
    bInit          : BOOL := FALSE;         // 首扫标志，初值 FALSE，判据 NOT bInit [-] / First-scan flag initialised FALSE
    ePhase         : E_DL_GapPhase := E_DL_GapPhase.eIdle;  // 内部相位，对外经 eState 输出 / Internal phase, exported as eState
    fMinUse        : REAL;                  // 生效的指令下限 [毫米]，已按大小关系归一 / Effective lower limit, normalised by magnitude
    fMaxUse        : REAL;                  // 生效的指令上限 [毫米]，已按大小关系归一 / Effective upper limit, normalised by magnitude
    fSpUse         : REAL;                  // 钳位后的目标辊距 [毫米] / Clamped target roller gap
    fTolUse        : REAL;                  // 生效的到位容差 [毫米]，负值取绝对值 / Effective tolerance, negative input taken as absolute
    fBlUse         : REAL;                  // 生效的背隙补偿量 [毫米]，已钳位 / Effective backlash compensation, clamped
    fApproachTarget : REAL;                 // 越程过半判据点 [毫米] / Half overshoot threshold of the approach phase
    fCmdCandidate  : REAL;                  // 指令候选值，钳位前中间量 [毫米] / Command candidate before clamping
    fDeviation     : REAL;                  // 本次残余偏差中间量 [毫米] / Residual deviation of this adjustment
    bInTol         : BOOL;                  // 本拍偏差在容差内且反馈有效 [-] / Flag, deviation inside tolerance with valid feedback
    bMoveRun       : BOOL;                  // 限时计时器输入，先算后调 [-] / Timeout timer input, computed before the call
    bMoveTimeout   : BOOL;                  // 限时到拍标志 [-] / Timeout flag of this cycle
    bTimeoutEnable : BOOL;                  // 是否启用限时监控 [-] / Flag, timeout monitoring enabled
    tMoveUse       : TIME;                  // 生效的限时值 [毫秒] / Effective timeout value
    bFeedbackLost  : BOOL;                  // 本拍反馈丢失（使能前提下）[-] / Flag, feedback lost while enabled
    bSpClamped     : BOOL;                  // 目标被钳位的标记 [-] / Flag, the target was clamped
    bBlClamped     : BOOL;                  // 背隙被钳位的标记 [-] / Flag, the backlash was clamped
    bArrived       : BOOL;                  // 本拍刚到位，供统计段使用 [-] / Flag, arrival happened in this cycle
    bStateIllegal  : BOOL;                  // 非法相位被兜底捕获 [-] / Flag, an illegal phase was captured
END_VAR
VAR CONSTANT
    DL_FLOAT_EPS     : REAL := 1.0E-6;      // 浮点判零容差 [无量纲] / Float epsilon for zero tests
    DL_APPROACH_SIGN : REAL := -1.0;        // 逼近方向符号，负向吃背隙 [无量纲] / Approach direction sign, negative eats the backlash
    DL_BACKLASH_MAX  : REAL := 1.0;         // 背隙补偿上限 [毫米]，防组态错值 / Backlash compensation upper bound
    DL_OVERSHOOT_RATIO : REAL := 0.5;       // 越程过半判据比例 [无量纲] / Half overshoot ratio of the approach phase
    DL_DEV_ALPHA     : REAL := 0.2;         // 偏差均值一阶低通系数 [无量纲] / First order low pass coefficient of the deviation average
    DL_CNT_MAX       : UDINT := 16#FFFF_FFFE;  // 计数饱和上限，防溢出回绕 [次] / Counter saturation limit
    DL_TIME_ZERO     : TIME := T#0MS;       // 时间零值基准 [毫秒] / Time zero reference
    DL_TIME_NEVER    : TIME := T#24H;       // 限时关闭时的占位时长 [毫秒] / Placeholder duration when timeout monitoring is off
END_VAR

(*------------------------------------------------------------------------------
 * 段 1｜沿检测无条件刷新（R7 红线）
 *      Edge detection refreshed unconditionally
 *-----------------------------------------------------------------------------*)
fbTrigReset(CLK := bReset);
fbTrigStart(CLK := bAdjustStart);

(*------------------------------------------------------------------------------
 * 段 2｜首扫初始化（R19 唯一合法范式）
 *      First-scan initialisation with the canonical R19 pattern
 *-----------------------------------------------------------------------------*)
IF NOT bInit THEN
    fGapCmd        := 0.0;                 // 指令初值：由上层在投运时给定安全位
    bAdjusting     := FALSE;
    bInPosition    := FALSE;
    fLastDeviation := 0.0;
    nAdjustCount   := 0;
    ePhase         := E_DL_GapPhase.eIdle;
    eState         := E_DL_GapPhase.eIdle;
    bError         := FALSE;
    bStateIllegal  := FALSE;
    stTrim.fDevAvg     := 0.0;             // 偏差均值初值为零
    stTrim.tLastMove   := DL_TIME_ZERO;    // 耗时初值为零
    stTrim.nOverTolCnt := 0;               // 超容差次数初值为零
    uErrorId       := 16#0000_0000;
    bInit          := TRUE;                // 首扫只做一次
END_IF

(*------------------------------------------------------------------------------
 * 段 3｜参数钳位（先归一上下限，再钳目标与背隙；越界只记信息级码）
 *      Parameter clamping, normalise the limits first, info level only
 *-----------------------------------------------------------------------------*)
bSpClamped := FALSE;
bBlClamped := FALSE;

IF fCmdMax < fCmdMin THEN
    fMinUse    := fCmdMax;                 // 上下限颠倒：自动换位，避免非法区间
    fMaxUse    := fCmdMin;
    bSpClamped := TRUE;                    // 记入参数越界信息码
ELSE
    fMinUse := fCmdMin;
    fMaxUse := fCmdMax;
END_IF

IF fGapSetpoint < fMinUse THEN
    fSpUse     := fMinUse;                 // 低于下限：钳到下限
    bSpClamped := TRUE;
ELSIF fGapSetpoint > fMaxUse THEN
    fSpUse     := fMaxUse;                 // 高于上限：钳到上限
    bSpClamped := TRUE;
ELSE
    fSpUse := fGapSetpoint;
END_IF

IF fGapTol >= 0.0 THEN
    fTolUse := fGapTol;                    // 容差非负：原样使用
ELSE
    fTolUse := ABS(fGapTol);               // 容差为负：按绝对值理解
    bSpClamped := TRUE;
END_IF

IF fBacklash < 0.0 THEN
    fBlUse     := 0.0;                     // 负背隙无物理意义：按不补偿处理
    bBlClamped := TRUE;
ELSIF fBacklash > DL_BACKLASH_MAX THEN
    fBlUse     := DL_BACKLASH_MAX;         // 超上限：钳到上限
    bBlClamped := TRUE;
ELSE
    fBlUse := fBacklash;
END_IF

(*------------------------------------------------------------------------------
 * 段 4｜到位判定与限时准备（判定条件与计时输入都在此处一次算清）
 *      In-position judgement and timeout preparation, computed once here
 *-----------------------------------------------------------------------------*)
fDeviation := fGapActual - fSpUse;
IF bFeedbackValid AND (ABS(fDeviation) <= fTolUse) THEN
    bInTol := TRUE;                        // 偏差入带且反馈可信才算到位
ELSE
    bInTol := FALSE;
END_IF

IF tMoveTimeout <= DL_TIME_ZERO THEN
    tMoveUse       := DL_TIME_NEVER;       // 零限时：关闭监控，避免立即误报
    bTimeoutEnable := FALSE;
ELSE
    tMoveUse       := tMoveTimeout;
    bTimeoutEnable := TRUE;
END_IF

bMoveRun := (ePhase = E_DL_GapPhase.eApproach) OR (ePhase = E_DL_GapPhase.eFine);
fbTonMove(IN := bMoveRun, PT := tMoveUse);
bMoveTimeout := bTimeoutEnable AND fbTonMove.Q;

IF bEnable AND (NOT bFeedbackValid) THEN
    bFeedbackLost := TRUE;                 // 使能状态下反馈无效：按丢失处理
ELSE
    bFeedbackLost := FALSE;
END_IF

bArrived := FALSE;                         // 到位单拍标志预清零

(*------------------------------------------------------------------------------
 * 段 5｜主状态机（ENUM 加 CASE，含 ELSE 兜底；每成员均有对应标签）
 *      Main state machine, one label per enumeration member plus a fallback
 *      指令只在跃迁拍写，其余拍不写，从而天然满足「故障时指令保持」
 *-----------------------------------------------------------------------------*)
CASE ePhase OF
    E_DL_GapPhase.eIdle:
        IF NOT bEnable THEN
            bInPosition := FALSE;          // 未使能：位置不可信，撤回到位标志
        ELSIF fbTrigStart.Q THEN
            bInPosition := FALSE;          // 每次调整都从「未到位」开始记账
            IF bFeedbackLost THEN
                ePhase := E_DL_GapPhase.eFault;        // 反馈无效不得启动，指令保持
            ELSE
                fCmdCandidate := fSpUse + DL_APPROACH_SIGN * fBlUse;
                fGapCmd       := LIMIT(fMinUse, fCmdCandidate, fMaxUse);  // 越程值再钳一次
                ePhase        := E_DL_GapPhase.eApproach;
            END_IF
        END_IF

    E_DL_GapPhase.eApproach:
        IF NOT bEnable THEN
            ePhase := E_DL_GapPhase.eIdle;
        ELSIF bFeedbackLost THEN
            ePhase := E_DL_GapPhase.eFault;            // 反馈丢失：转故障，指令保持
        ELSIF bMoveTimeout THEN
            ePhase := E_DL_GapPhase.eFault;            // 越程段超时：转故障
        ELSE
            fApproachTarget := fSpUse + DL_APPROACH_SIGN * fBlUse * DL_OVERSHOOT_RATIO;
            IF (DL_APPROACH_SIGN * (fGapActual - fApproachTarget)) >= 0.0 THEN
                fGapCmd := LIMIT(fMinUse, fSpUse, fMaxUse);   // 越程过半：回目标值
                ePhase  := E_DL_GapPhase.eFine;
            END_IF
        END_IF

    E_DL_GapPhase.eFine:
        IF NOT bEnable THEN
            ePhase := E_DL_GapPhase.eIdle;
        ELSIF bFeedbackLost THEN
            ePhase := E_DL_GapPhase.eFault;            // 反馈丢失：转故障，指令保持
        ELSIF bInTol THEN
            fGapCmd        := LIMIT(fMinUse, fSpUse, fMaxUse);   // 到位拍指令即目标值
            fLastDeviation := fDeviation;              // 残余偏差：带符号，正为偏大
            bInPosition    := TRUE;
            bArrived       := TRUE;                    // 供统计段使用
            ePhase         := E_DL_GapPhase.eHold;
        ELSIF bMoveTimeout THEN
            ePhase := E_DL_GapPhase.eFault;            // 精定位超时：转故障
        END_IF

    E_DL_GapPhase.eHold:
        IF NOT bEnable THEN
            bInPosition := FALSE;                      // 未使能撤回到位标志
            ePhase      := E_DL_GapPhase.eIdle;
        ELSIF fbTrigStart.Q THEN
            bInPosition := FALSE;                      // 新一轮调整：先撤到位
            IF bFeedbackLost THEN
                ePhase := E_DL_GapPhase.eFault;
            ELSE
                fCmdCandidate := fSpUse + DL_APPROACH_SIGN * fBlUse;
                fGapCmd       := LIMIT(fMinUse, fCmdCandidate, fMaxUse);
                ePhase        := E_DL_GapPhase.eApproach;
            END_IF
        ELSIF bFeedbackLost THEN
            bInPosition := FALSE;                      // 位置不可信：撤回到位，但不断开保持
            ePhase      := E_DL_GapPhase.eFault;
        END_IF

    E_DL_GapPhase.eFault:
        IF NOT bEnable THEN
            ePhase := E_DL_GapPhase.eIdle;             // 停使能可直接退出故障态
        ELSIF fbTrigReset.Q THEN
            ePhase        := E_DL_GapPhase.eIdle;      // 复位后回待机，指令保持原值
            bStateIllegal := FALSE;
        END_IF

    ELSE
        ePhase        := E_DL_GapPhase.eFault;         // 非法值兜底
        bStateIllegal := TRUE;
END_CASE

(*------------------------------------------------------------------------------
 * 段 6｜统计记账（只在到位拍更新，避免逐拍累加污染台账）
 *      Statistics updated on the arrival cycle only
 *-----------------------------------------------------------------------------*)
IF bArrived THEN
    IF ABS(stTrim.fDevAvg) < DL_FLOAT_EPS THEN
        stTrim.fDevAvg := fLastDeviation;              // 首次到位：均值直接取本次值
    ELSE
        stTrim.fDevAvg := stTrim.fDevAvg + DL_DEV_ALPHA * (fLastDeviation - stTrim.fDevAvg);
    END_IF
    stTrim.tLastMove := fbTonMove.ET;                  // 本次耗时取限时器已计时间
    IF ABS(fLastDeviation) > fTolUse THEN
        IF stTrim.nOverTolCnt < DL_CNT_MAX THEN
            stTrim.nOverTolCnt := stTrim.nOverTolCnt + 1;
        END_IF
    END_IF
    IF nAdjustCount < DL_CNT_MAX THEN
        nAdjustCount := nAdjustCount + 1;               // 仅到位才计入次数
    END_IF
END_IF

(*------------------------------------------------------------------------------
 * 段 7｜输出归并与码位定级（单一优先级链，全拍只写一次 uErrorId）
 *      Output merge and single-priority error code resolution
 *-----------------------------------------------------------------------------*)
bAdjusting := (ePhase = E_DL_GapPhase.eApproach) OR (ePhase = E_DL_GapPhase.eFine);

IF bStateIllegal THEN
    uErrorId := 16#0003_0308;                          // 优先级一：非法相位
ELSIF bFeedbackLost THEN
    uErrorId := 16#0003_0306;                          // 优先级二：反馈无效或丢失
ELSIF bMoveTimeout THEN
    uErrorId := 16#0003_0305;                          // 优先级三：到位超时
ELSIF bSpClamped THEN
    uErrorId := 16#0003_0147;                          // 信息级：目标越界已钳位
ELSIF bBlClamped THEN
    uErrorId := 16#0003_0148;                          // 信息级：背隙越界已钳位
ELSE
    uErrorId := 16#0000_0000;
END_IF

(* 故障位只反映故障级：信息级码 0147 与 0148 绝不置故障位（R21） *)
bError := bStateIllegal OR bFeedbackLost OR bMoveTimeout;

eState := ePhase;                                      // 相位每拍重写，供 HMI 诊断
END_FUNCTION_BLOCK
